(* IEC 61131-3 sources: daoli-st-library/DL_Device (part 21) *)

(* ---- FB_DL_EscChuckCurrentMonitor.st ---- *)
(*
    FB_DL_EscChuckCurrentMonitor —— ESC 静电吸附电流监视
    ------------------------------------------------------------------
    分类      : DL_Device / Diagnostics
    前缀      : FB_DL_
    版本      : 1.0.0
    溯源      : 半导体静电吸盘（ESC）自研线，clean-room 自研，无可挖开源源；
                只借公开半导体设备工程语义（吸附/建立/稳态/释放三段，失吸与打火是
                可区分的失效模式）；判据、状态机、错误分级与码位 100% 自有；
                E_DL_Ne107Status 属主为 I_DL_DeviceHealth，本件只引用不重声明（R70）
    平台      : 纯 IEC 61131-3，CODESYS V3.5+ / TwinCAT 3 / InoProShop 通用
    作者      : 道莅代码库 · PLC编程专家（R19）
    ------------------------------------------------------------------
    功能说明  : 吸附电压施加后电流须在 tBuildTime 内落进电流窗（建立段）；之后电流须
                持续落窗（稳态段，低于下限超 tConfirmTime 判失吸）；撤电压后电流须归零
                （释放段）。失吸会导致晶圆飞片/破片，打火会烧盘面，两者在电流波形上
                是两种截然不同的特征，本件把「电流长时间偏低」与「瞬时尖峰」分开判。
                核心防御：① 阈值倒置先自动交换并置信息码，交换后仍非法才报故障级；
                ② 电流/电压非有限即故障级并冻结判定，且保持末次 bAttached——
                   把正在吸附的晶圆判成飞片会引发误停机；
                ③ 电压低于吸附门限时不判电流（电压没加上，电流当然为零），回 eIdle；
                ④ 打火只锁存并出口 eOutOfSpec，不置 bError（可继续生产但需检修）；
                ⑤ 泄漏趋势用前后半窗均值比较，只置信息级不置故障。
                职责边界：吸附电压给定与放电归静电电源件，本件只判电流形态。
    错误码    : 16#0003_016E 电流窗上下限倒置已自动交换 / 泄漏趋势上升 / 贴近边界降级运行——信息级，正常防御
                16#0003_016F 预留禁用（信息级，不得挪用）
                16#0003_0336 阈值参数非法或输入非有限——故障级，判定冻结且保持末次吸附结论
                16#0003_0337 建立超时或稳态电流失窗（判失吸）——故障级，eHealth = eFailure
                16#0003_0338 打火尖峰锁存——故障级码位且 eHealth = eOutOfSpec，但按 R13 家族裁定不置 bError
    码位总账  : 16#0003_016E 用 / 16#0003_016F 预留 ｜ 16#0003_0336 用 / 16#0003_0337 用 / 16#0003_0338 用
    状态机    : E_DL_EscState（eIdle / eBuild / eSteady / eRelease / eFault）五态，CASE 含 ELSE 兜底，
                ELSE 回 eFault 并置故障级 0336。
    采样约定  : fbTrigReset / fbBuild / fbLossConfirm 在本体首部无条件刷新——两个定时器的 IN
                由状态导出但调用绝不放进 IF 或 CASE（按段断输入是本族高危点）；
                采样周期越域即故障级，因为趋势窗与确认时间都隐含依赖采样节拍。
    修订记录  : 2026-11-16 v1.0.0 首次入库（R19）
*)

(*
    枚举 : E_DL_EscState —— 静电吸盘工作段（本文件为全库唯一属主）
*)
TYPE E_DL_EscState :
(
    eIdle    := 0,                            // 空闲：未施加吸附电压 / idle, no chuck voltage applied
    eBuild   := 1,                            // 建立段：等待电流落窗 / build phase, waiting for the current to settle
    eSteady  := 2,                            // 稳态段：电流持续落窗 / steady phase, the current stays inside the window
    eRelease := 3,                            // 释放段：等待电流归零 / release phase, waiting for the current to vanish
    eFault   := 4                             // 故障：判定冻结 / fault, evaluation frozen
);
END_TYPE

FUNCTION_BLOCK FB_DL_EscChuckCurrentMonitor
VAR_INPUT
    bEnable         : BOOL;                   // 使能，FALSE 撤销所有判定输出 / enable, FALSE withdraws every judgement output
    bReset          : BOOL;                   // 复位，上升沿清故障与趋势 / reset, rising edge clears the faults and the trend
    bChuckOn        : BOOL := FALSE;          // 吸附电压施加命令（上层给定）/ chuck voltage command from the upper layer
    fChuckCurrent   : REAL := 0.0;            // 吸附电流测量值 [uA]，范围 0.0~10000.0 / chuck current measurement [uA], range 0.0~10000.0
    fChuckVoltage   : REAL := 0.0;            // 吸附电压测量值 [V]，范围 0.0~5000.0 / chuck voltage measurement [V], range 0.0~5000.0
    fCurMin         : REAL := 5.0;            // 稳态电流窗下限 [uA]，必须 > 0 / steady window lower bound [uA], must be > 0
    fCurMax         : REAL := 500.0;          // 稳态电流窗上限 [uA]，必须 > fCurMin / steady window upper bound [uA], must be > fCurMin
    fSparkRise      : REAL := 50.0;           // 打火判据：单拍电流跳变量阈值 [uA]，必须 > 0 / spark criterion, per cycle current step [uA], must be > 0
    tBuildTime      : TIME := T#2S;           // 建立段允许时长 [ms]，范围 100~30000 / build phase allowance [ms], range 100~30000
    tConfirmTime    : TIME := T#500MS;        // 失吸确认时间 [ms]，范围 0~10000 / loss confirmation time [ms], range 0~10000
    tSampleTime     : TIME := T#10MS;         // 采样周期 [ms]，范围 1~1000 / sample time [ms], range 1~1000
END_VAR
VAR_OUTPUT
    bAttached       : BOOL;                   // 判定已吸附（建立成功且稳态落窗）/ attached, build succeeded and the steady current stays in the window
    bSpark          : BOOL;                   // 检出打火尖峰（锁存）/ spark peak detected, latched
    bLeakTrend      : BOOL;                   // 泄漏趋势上升（盘面污染或绝缘退化）/ leakage trend rising, contamination or insulation ageing
    bDegraded       : BOOL;                   // 降级运行（电流在窗内但贴近边界）/ degraded, the current is in the window but close to a bound
    eHealth         : E_DL_Ne107Status;       // 健康出口（引用唯一属主枚举）/ health output referencing the owner enumeration
    uAttachCount    : UDINT;                  // 累计成功吸附次数，饱和 [次] / accumulated successful attaches, saturating [times]
    eErr            : UDINT;                  // 错误码，0=正常 / error id, 0=ok
    bError          : BOOL;                   // 故障标志，eErr 为故障级时 TRUE / error flag, TRUE on fault-level eErr
END_VAR
VAR
    eState          : E_DL_EscState := eIdle; // 状态机当前态 / current state machine state
    fbTrigReset     : R_TRIG;                 // 复位上升沿实例，本体首部无条件刷新 / reset edge instance, refreshed unconditionally
    fbBuild         : TON;                    // 建立段定时器，本体首部无条件刷新 / build phase timer, refreshed unconditionally
    fbLossConfirm   : TON;                    // 失吸确认定时器，本体首部无条件刷新 / loss confirmation timer, refreshed unconditionally
    fPrevCur        : REAL;                   // 上一拍电流，用于打火跳变判据 [uA] / previous current for the spark step test [uA]
    fTrendAcc       : REAL;                   // 后窗电流均值累加 [uA] / second window current mean accumulator [uA]
    fTrendBase      : REAL;                   // 前窗电流均值累加 [uA] / first window current mean accumulator [uA]
    uTrendCnt       : UINT;                   // 趋势取样计数 [拍] / trend sampling counter [scan]
    fCurMinEff      : REAL;                   // 交换与钳位后的电流窗下限 [uA] / effective lower bound after swap and clamp [uA]
    fCurMaxEff      : REAL;                   // 交换与钳位后的电流窗上限 [uA] / effective upper bound after swap and clamp [uA]
    fBandEff        : REAL;                   // 近边界判定带宽 [uA] / near boundary band width [uA]
    fCur            : REAL;                   // 本拍电流副本 [uA] / current copy of this cycle [uA]
    bNonFin         : BOOL;                   // 输入非有限判定标志 / non-finite input flag
    bInWindow       : BOOL;                   // 电流落窗判定 / current inside the window
    bInit           : BOOL := FALSE;          // 首扫标志，初值 FALSE，判据 NOT bInit / first-scan flag, initial FALSE, tested with NOT
END_VAR
VAR CONSTANT
    DL_ESC_CUR_ABS_MAX : REAL := 10000.0;     // 电流绝对上限（三阈值钳位用）[uA] / absolute current bound used by the clamps [uA]
    DL_ESC_VOLT_MIN    : REAL := 100.0;       // 判定「电压确实加上了」的下限 [V] / lower bound proving the voltage is really applied [V]
    DL_ESC_TREND_N     : UINT := 50;          // 趋势取样个数 [拍] / number of trend samples [scan]
    DL_ESC_BAND_RATIO  : REAL := 0.05;        // 近边界判定带宽（相对窗宽）[无量纲] / near boundary band relative to the window [dimensionless]
    DL_ESC_DT_MAX      : TIME := T#1S;        // 采样周期上限 [ms] / sample time upper bound [ms]
    DL_ESC_DT_MIN      : TIME := T#1MS;       // 采样周期下限 [ms] / sample time lower bound [ms]
    DL_FLOAT_EPS       : REAL := 1.0E-6;      // 浮点判等容差 [无量纲] / float equality tolerance [dimensionless]
    DL_ESC_TWO         : REAL := 2.0;         // 二值常量，窗口折半用 [无量纲] / two, used to halve the trend window
    DL_ESC_INF_GUARD   : REAL := 1.0E38;      // 非有限幅值判定阈值 [无量纲] / non-finite magnitude guard [dimensionless]
    DL_ESC_CNT_MAX     : UDINT := 16#FFFF_FFFE; // 吸附计数饱和值 [次] / attach counter saturation value [times]
    DL_ESC_ZERO        : REAL := 0.0;         // 零值常量，避免裸字面量 [无量纲] / zero constant, avoids a bare literal [dimensionless]
END_VAR

// 段 1｜边沿与定时器实例无条件周期刷新（红线：严禁放入条件分支）/ segment 1, unconditional refresh
fbTrigReset(CLK := bReset);
fbBuild(IN := (eState = eBuild) AND bEnable, PT := tBuildTime); // 仅建立段计时 / the timer runs only during the build phase
fbLossConfirm(IN := (eState = eSteady) AND bEnable AND (fChuckCurrent < fCurMin), PT := tConfirmTime); // 仅稳态且电流低于下限时计时 / runs only in the steady phase while the current is below the bound

// 段 2｜输出与错误状态预置（bAttached / bSpark 为保持量，不预置）/ segment 2, preset outputs, the held flags are not preset
eErr := 0;                                    // 预置无错误 / preset no error
bError := FALSE;                              // 预置无故障 / preset no fault
bDegraded := FALSE;                           // 预置未降级 / preset not degraded
bLeakTrend := FALSE;                          // 预置无泄漏趋势 / preset no leakage trend
eHealth := eOk;                               // 预置健康 / preset OK

// 段 3｜首扫初始化（唯一合法范式：初值 FALSE，判据 NOT bInit）/ segment 3, first-scan initialisation
IF NOT bInit THEN
    bAttached := FALSE;                       // 首扫不判吸附 / no attach survives the first scan
    bSpark := FALSE;                          // 首扫不打火锁存 / no spark latch survives the first scan
    uAttachCount := 0;                        // 吸附计数清零 / clear the attach counter
    fPrevCur := fChuckCurrent;                // 电流基准取当前测量，避免首拍误判打火 / seed the current reference to avoid a false spark on the first scan
    uTrendCnt := 0;                          // 趋势计数清零 / clear the trend counter
    fTrendAcc := DL_ESC_ZERO;                 // 后窗累加清零 / clear the second window accumulator
    fTrendBase := DL_ESC_ZERO;                // 前窗累加清零 / clear the first window accumulator
    bInit := TRUE;                            // 首扫只做一次 / first scan runs once only
END_IF

// 段 4｜使能闸：失能撤销全部判定输出 / segment 4, enable gate
IF NOT bEnable THEN
    bAttached := FALSE;                       // 撤销吸附判定 / withdraw the attach judgement
    bDegraded := FALSE;                       // 撤销降级 / withdraw the degraded flag
    bLeakTrend := FALSE;                      // 撤销趋势 / withdraw the trend flag
    eHealth := eUnknown;                      // 失能即未知 / unknown while disabled
    RETURN;                                   // 失能即出口 / disabled is the exit
END_IF

// 段 5｜阈值交换与合法性闸（倒置先交换，交换后仍非法才报故障）/ segment 5, threshold swap and validity
fCurMinEff := fCurMin;                        // 取入参副本 / copy the input
fCurMaxEff := fCurMax;                        // 取入参副本 / copy the input
IF fCurMaxEff < fCurMinEff THEN
    fCurMinEff := fCurMax;                    // 交换：下限取原上限 / swap, the lower bound takes the former upper bound
    fCurMaxEff := fCurMin;                    // 交换：上限取原下限 / swap, the upper bound takes the former lower bound
    eErr := 16#0003_016E;                     // 信息级：上下限倒置已自动交换 / info level, the inverted bounds were swapped
END_IF
fCurMinEff := MIN(MAX(fCurMinEff, DL_ESC_ZERO), DL_ESC_CUR_ABS_MAX); // 下限收敛到物理域 / converge the lower bound into the physical domain
fCurMaxEff := MIN(MAX(fCurMaxEff, DL_ESC_ZERO), DL_ESC_CUR_ABS_MAX); // 上限收敛到物理域 / converge the upper bound into the physical domain
IF (fCurMinEff <= DL_FLOAT_EPS) OR (fCurMaxEff <= fCurMinEff) THEN
    eErr := 16#0003_0336;                     // 阈值非法故障码 / illegal threshold fault id
    bError := TRUE;                           // 置故障标志 / raise the error flag
    eState := eFault;                         // 落故障态，判定冻结 / enter the fault state, the evaluation is frozen
    eHealth := eFailure;                      // 阈值不可信即出口失效 / untrustworthy thresholds mean a failed health output
    RETURN;                                   // 故障级提前返回，bAttached 保持末值 / early return, bAttached keeps its last value
END_IF
fBandEff := DL_ESC_BAND_RATIO * (fCurMaxEff - fCurMinEff); // 近边界带宽 [uA] / near boundary band width [uA]

// 段 6｜输入非有限闸：冻结判定并保持末次吸附结论 / segment 6, non-finite gate freezes the judgement
bNonFin := (fChuckCurrent <> fChuckCurrent) OR (fChuckCurrent > DL_ESC_INF_GUARD) OR (fChuckCurrent < -DL_ESC_INF_GUARD)
        OR (fChuckVoltage <> fChuckVoltage) OR (fChuckVoltage > DL_ESC_INF_GUARD) OR (fChuckVoltage < -DL_ESC_INF_GUARD)
        OR (fSparkRise <> fSparkRise);        // 非有限判定 / non-finite detection
IF bNonFin THEN
    eErr := 16#0003_0336;                     // 输入非有限故障码 / non-finite input fault id
    bError := TRUE;                           // 置故障标志 / raise the error flag
    eState := eFault;                         // 落故障态 / enter the fault state
    eHealth := eFailure;                      // 测量不可信 / the measurement is untrustworthy
    RETURN;                                   // 保持末次 bAttached，绝不掉成未吸附 / keep the last attach state, never fall back to detached
END_IF

// 段 7｜采样周期闸（趋势窗与确认时间都依赖采样节拍）/ segment 7, sample time gate
IF (tSampleTime < DL_ESC_DT_MIN) OR (tSampleTime > DL_ESC_DT_MAX) THEN
    eErr := 16#0003_0336;                     // 采样周期非法故障码 / illegal sample time fault id
    bError := TRUE;                           // 置故障标志 / raise the error flag
    eState := eFault;                         // 落故障态 / enter the fault state
    eHealth := eFailure;                      // 节拍不可信 / the timing is untrustworthy
    RETURN;                                   // 出口 / exit
END_IF

// 段 8｜复位沿清故障与趋势（不改变已建立的吸附结论）/ segment 8, reset clears the faults and the trend
IF fbTrigReset.Q THEN
    bSpark := FALSE;                          // 清打火锁存 / clear the spark latch
    bLeakTrend := FALSE;                      // 清趋势 / clear the trend
    uTrendCnt := 0;                           // 清趋势计数 / clear the trend counter
    fTrendAcc := DL_ESC_ZERO;                 // 清后窗累加 / clear the second window
    fTrendBase := DL_ESC_ZERO;                // 清前窗累加 / clear the first window
    IF eState = eFault THEN
        eState := eIdle;                      // 故障态复位回空闲 / a reset leaves the fault state
    END_IF
END_IF

// 段 9｜电流副本与落窗判定 / segment 9, current copy and window test
fCur := fChuckCurrent;                        // 取入参副本 [uA] / copy the input [uA]
bInWindow := (fCur >= fCurMinEff) AND (fCur <= fCurMaxEff); // 落窗判定 / window test

// 段 10｜打火判据（单拍跳变 + 吸附电压在场，只锁存不置 bError）/ segment 10, spark criterion
IF bChuckOn AND (ABS(fCur - fPrevCur) > fSparkRise) THEN
    bSpark := TRUE;                           // 锁存打火 / latch the spark
    eErr := 16#0003_0338;                     // 打火故障级码位，但按家族裁定不置 bError / spark fault id without raising bError
    eHealth := eOutOfSpec;                    // 能继续吸不等于盘面完好 / still holding does not mean the chuck surface is intact
END_IF
fPrevCur := fCur;                             // 记录本拍电流供下一拍比较 / remember this cycle current

// 段 11｜降级判定：电流在窗内但贴近上下边界 / segment 11, degraded evaluation near a bound
IF bInWindow AND ((fCur <= (fCurMinEff + fBandEff)) OR (fCur >= (fCurMaxEff - fBandEff))) THEN
    bDegraded := TRUE;                        // 贴近边界即降级 / closeness to a bound is a degradation
    IF eErr = 0 THEN
        eErr := 16#0003_016E;                 // 信息级：贴近边界降级运行 / info level, running degraded near a bound
    END_IF
END_IF

// 段 12｜泄漏趋势（前后半窗均值比较，只置信息级）/ segment 12, leakage trend by half window means
IF eState = eSteady THEN
    IF uTrendCnt < (DL_ESC_TREND_N / 2) THEN
        fTrendBase := fTrendBase + fCur / (UINT_TO_REAL(DL_ESC_TREND_N) / DL_ESC_TWO); // 前窗均值累加 [uA] / accumulate the first window mean [uA]
        uTrendCnt := uTrendCnt + 1;           // 计数加一 / increment the counter
    ELSE
        fTrendAcc := fTrendAcc + fCur / (UINT_TO_REAL(DL_ESC_TREND_N) / DL_ESC_TWO);   // 后窗均值累加 [uA] / accumulate the second window mean [uA]
        uTrendCnt := uTrendCnt + 1;           // 计数加一 / increment the counter
        IF uTrendCnt >= DL_ESC_TREND_N THEN
            IF fTrendAcc > (fTrendBase + DL_ESC_BAND_RATIO * (fCurMaxEff - fCurMinEff)) THEN
                bLeakTrend := TRUE;           // 后窗显著上爬：污染或绝缘退化 / the second window creeps up, contamination or insulation ageing
                eErr := 16#0003_016E;         // 信息级：泄漏趋势上升 / info level, the leakage trend is rising
                eHealth := eMaintenanceReq;   // 需安排检修 / maintenance is required
            END_IF
            uTrendCnt := 0;                   // 窗口滑动复位 / restart the sliding window
            fTrendAcc := DL_ESC_ZERO;         // 后窗累加清零 / clear the second window
            fTrendBase := DL_ESC_ZERO;        // 前窗累加清零 / clear the first window
        END_IF
    END_IF
END_IF

// 段 13｜状态机（含 ELSE 兜底）/ segment 13, state machine with ELSE fallback
CASE eState OF
    eIdle:
        bAttached := FALSE;                   // 空闲即未吸附 / idle means detached
        IF bChuckOn AND (fChuckVoltage >= DL_ESC_VOLT_MIN) THEN
            eState := eBuild;                 // 电压确实加上才进入建立段 / enter the build phase only when the voltage is really present
        END_IF

    eBuild:
        IF bInWindow THEN
            eState := eSteady;                // 电流落窗即建立成功 / the current entering the window completes the build
            bAttached := TRUE;                // 判定已吸附 / mark it attached
            IF uAttachCount < DL_ESC_CNT_MAX THEN
                uAttachCount := uAttachCount + 1; // 饱和计数 / saturating count
            END_IF
        ELSIF fbBuild.Q THEN
            eErr := 16#0003_0337;             // 建立超时故障码 / build timeout fault id
            bError := TRUE;                   // 置故障标志 / raise the error flag
            eHealth := eFailure;              // 失吸 / the wafer is not held
            eState := eFault;                 // 落故障态 / enter the fault state
            bAttached := FALSE;               // 建立失败即未吸附 / a failed build means detached
        END_IF

    eSteady:
        bAttached := TRUE;                    // 稳态保持吸附 / the steady phase keeps the attach state
        IF NOT bChuckOn THEN
            eState := eRelease;               // 撤电压即进入释放段 / releasing the voltage enters the release phase
        ELSIF fbLossConfirm.Q THEN
            eErr := 16#0003_0337;             // 失吸确认故障码 / loss confirmation fault id
            bError := TRUE;                   // 置故障标志 / raise the error flag
            eHealth := eFailure;              // 失吸 / the wafer is lost
            eState := eFault;                 // 落故障态 / enter the fault state
            bAttached := FALSE;               // 确认失吸 / confirmed detached
        END_IF

    eRelease:
        bAttached := FALSE;                   // 释放段即不再算吸附 / the release phase is not an attached state
        IF fCur <= DL_FLOAT_EPS THEN
            eState := eIdle;                  // 电流归零即回空闲 / back to idle once the current vanishes
        ELSIF bChuckOn THEN
            eState := eBuild;                 // 释放过程中重新上电：重新建立 / re-energising during release restarts the build
        END_IF

    eFault:
        bAttached := FALSE;                   // 故障态不判吸附 / no attach judgement in the fault state
        IF NOT bChuckOn THEN
            eState := eIdle;                  // 撤电压允许退出故障态（复位亦可）/ withdrawing the voltage also leaves the fault state
        END_IF

ELSE
    eErr := 16#0003_0336;                     // 故障级：非法状态兜底 / fault level, illegal state fallback
    bError := TRUE;                           // 置故障标志 / raise the error flag
    eState := eFault;                         // 回故障态 / fall back to the fault state
    eHealth := eUnknown;                      // 状态不可信 / the state is untrustworthy
END_CASE
END_FUNCTION_BLOCK

(* ---- FB_DL_EsdGroundMonitor.st ---- *)
(*
  ==================================================================
  组件名 Component  : FB_DL_EsdGroundMonitor
  分类   Category   : DL_Device
  复杂度 Complexity  : cx4
  版本   Version    : 1.0.0
  功能   Purpose    : ESD 接地连续性监视。对接地电阻做窗口判级（低于下限疑短路 /
                      接线反，高于上限疑断路），双阈值迟滞防边界抖动；传感失效
                      锁存优先于判级；健康语言出口按 NE107 五态口径输出。
  来源   Source     : self-esc（次源 t2-8 NE107，借鉴 NE107 健康状态五态语言，
                      clean-room 自研实现，未复制任何文档代码行）
  溯源   Origin     : IEC 61131-3 标准语义的道莅防御性实现；ESD 接地电阻窗口
                      判级为公开防静电工艺语义（常见口径 <10 欧姆量级）。
  平台   Platform   : 纯 IEC 61131-3（LREAL 运算，无私有库、无定时器实例）
  分工声明 Split     : 与 DL_Device 存量联锁族（风机关 / 传递窗）分工——本件只
                      做接地电阻判级与健康语言映射，不做风量联锁与顺控。
  作者   Author     : 道莅代码库 · PLC 编程专家（R57）
  ------------------------------------------------------------------
  边界 Boundary     :
                      一 组态闸（R151）：fOhmMin > 0 且 fOhmMax > fOhmMin，
                         迟滞带宽 0 <= fHystOhm < 半窗宽；
                      二 迟滞收窄口径：进入判据用全带宽，退出判据带宽收窄
                         fHystOhm，防边界抖动反复置清；
                      三 传感失效（非有限双判据 / 电阻 < 0）锁存优先于判级；
                      四 成因锁存解除路径 = bReset 上升沿（唯一路径，R188）；
                      五 无全局变量、无外部变量声明、无物理地址寻址。
  输出契约 Output contract:
                      eHealth 为 NE107 五态健康语言；bGroundOk 为放行派生电平；
                      eFault 为锁存回放；bError 与故障级成因配对（R45）。
  修订记录 Revision  :
    2026-11-21  v1.0.0  R57 首版（批 4 · 序号 16）
  ==================================================================
*)

TYPE E_DL_EgmPhase :
(
    eIdle  := 0,  // 未使能：判级停摆 / disabled, the grading idle
    eRun   := 10, // 运行：逐拍判级 / running, graded every scan
    eFault := 90  // 故障：成因锁存 / fault, the cause latched
);
END_TYPE

TYPE E_DL_EgmFault :
(
    eNone       := 0, // 无成因 / no cause
    eCfgIllegal := 1, // 组态非法：电阻窗或迟滞越域（故障级，与 bError 配对）/ an illegal config
    eSensorBad  := 2, // 传感失效：电阻非有限或负值（故障级，与 bError 配对）/ a sensor failure
    eGroundOpen := 3, // 接地断路：电阻超上限（故障级，与 bError 配对）/ a ground open
    eGroundShort:= 4, // 接地短路疑点：电阻低于下限（故障级，与 bError 配对）/ a ground short suspect
    ePhaseBad   := 5  // 非法相位兜底（故障级，与 bError 配对）/ an illegal phase fallback
);
END_TYPE

TYPE E_DL_EgmHealth :
(
    eInit           := 0, // NE107 初始态 / the NE107 initial state
    eGood           := 1, // NE107 正常 / the NE107 good state
    eCheckFunction  := 2, // NE107 功能受影响（组态非法驻留）/ the NE107 check function state
    eMaintenanceReq := 3, // NE107 维护要求（判级异常驻留）/ the NE107 maintenance required state
    eFailure        := 4  // NE107 故障（传感失效锁存）/ the NE107 failure state
);
END_TYPE

FUNCTION_BLOCK FB_DL_EsdGroundMonitor
VAR_INPUT
    bEnable   : BOOL := TRUE;   // 使能，失能时判级停摆 [-] / enable, the grading stops when disabled
    bReset    : BOOL := FALSE;  // 复位上升沿清全部成因锁存 [-] / reset rising edge clears every cause latch
    fResOhm   : LREAL := 5.0;   // 接地电阻实测 [欧姆] / the measured ground resistance [ohm]
    fOhmMin   : LREAL := 0.5;   // 电阻窗下限 [欧姆]，域 大于零 / the window floor [ohm], above zero
    fOhmMax   : LREAL := 10.0;  // 电阻窗上限 [欧姆]，域 大于下限 / the window ceiling [ohm], above the floor
    fHystOhm  : LREAL := 0.5;   // 迟滞带宽 [欧姆]，域 0..半窗宽 / the hysteresis band [ohm]
END_VAR
VAR_OUTPUT
    eHealth  : E_DL_EgmHealth := E_DL_EgmHealth.eInit; // NE107 健康语言出口 [枚举] / the NE107 health outlet [enum]
    bGroundOk: BOOL := FALSE; // 接地合格放行派生电平 [-] / the ground ok derived level
    ePhase   : E_DL_EgmPhase := E_DL_EgmPhase.eIdle; // 相位出口 [枚举] / the phase outlet [enum]
    eFault   : E_DL_EgmFault := E_DL_EgmFault.eNone; // 成因出口，锁存回放 [枚举] / the cause outlet replayed from the latch
    bError   : BOOL := FALSE; // 故障锁存标志 [-] / the fault latch flag
END_VAR
VAR
    rtReset : R_TRIG; // 复位沿检测，段 0 无条件刷新 / the reset edge, refreshed unconditionally
    _ePhase : E_DL_EgmPhase := E_DL_EgmPhase.eIdle; // 内部相位，CASE 唯一写入目标 / the internal phase
    _eFaulC : E_DL_EgmFault := E_DL_EgmFault.eNone; // 故障级成因，锁存至复位沿 / the fault cause, latched until the reset edge
    _bFault : BOOL := FALSE; // 故障锁存位 [-] / the fault latch bit
    _bInit  : BOOL := FALSE; // 首扫初始化完成标志（R310）/ the first scan flag
    _bInOk  : BOOL := FALSE; // 电阻有限且非负 [-] / the resistance finite and nonnegative
    _bCfgOk : BOOL := FALSE; // 组态域内 [-] / the configuration inside the domain
    _bOpen  : BOOL := FALSE; // 断路迟滞锁存 [-] / the open hysteresis latch
    _bShort : BOOL := FALSE; // 短路疑点迟滞锁存 [-] / the short suspect hysteresis latch
END_VAR

// 段 0｜沿检测无条件周期刷新（禁入分支）/ segment 0, the unconditional refresh
rtReset(CLK := bReset); // 复位沿 / the reset edge

// 段 1｜首扫初始化（R310）/ segment 1, the first scan initialisation
IF NOT _bInit THEN // 首扫一拍 / the first scan
    _bInit  := TRUE; // 置首扫标志 / raise the flag
    _ePhase := E_DL_EgmPhase.eRun; // 相位从运行起步（使能默认真）/ the phase starts in run
END_IF

// 段 2｜复位沿作用域：清锁存 / 清迟滞 / 迁相位（三项逐项声明）/ segment 2, the reset edge scope
IF rtReset.Q THEN // 复位沿 / the reset edge
    _bFault := FALSE; // 作用域一：清故障锁存 / scope one, clear the fault latch
    _eFaulC := E_DL_EgmFault.eNone; // 作用域一：清成因 / scope one, clear the cause
    _bOpen := FALSE; // 作用域二：清断路迟滞 / scope two, clear the open latch
    _bShort := FALSE; // 作用域二：清短路迟滞 / scope two, clear the short latch
    _ePhase := E_DL_EgmPhase.eRun; // 作用域三：迁回运行相 / scope three, back to run
END_IF

// 段 3｜组态与输入域闸（R151 全覆盖，边界一）/ segment 3, the configuration and input gates
_bInOk := (fResOhm = fResOhm) AND ((fResOhm - fResOhm) = (fResOhm - fResOhm)) AND (fResOhm >= 0.0); // 电阻有限且非负 / the resistance finite and nonnegative
_bCfgOk := (fOhmMin > 0.0) AND (fOhmMin = fOhmMin) AND (fOhmMax > fOhmMin) AND (fOhmMax = fOhmMax) AND (fHystOhm >= 0.0) AND (fHystOhm < (fOhmMax - fOhmMin) / 2.0); // 窗与迟滞域判定（除子为窗宽已证大于零）/ the window and hysteresis verdict
IF (NOT _bInOk) OR (NOT _bCfgOk) THEN // 输入缺陷或组态非法 / an input defect or an illegal config
    IF NOT _bFault THEN // 未锁存才迁移（防同拍抹除）/ migrate only while unlatched
        _bFault := TRUE; // 置故障锁存 / raise the fault latch
        IF NOT _bInOk THEN // 传感失效优先归因（R190 归因唯一）/ the sensor failure attributed first
            _eFaulC := E_DL_EgmFault.eSensorBad; // 传感失效成因 / the sensor cause
        ELSE // 组态非法 / the illegal config
            _eFaulC := E_DL_EgmFault.eCfgIllegal; // 组态成因 / the config cause
        END_IF
        _ePhase := E_DL_EgmPhase.eFault; // 迁故障相 / migrate to fault
    END_IF
END_IF

// 段 4｜相位机：ENUM + CASE，含 ELSE 非法相位兜底（R128）/ segment 4, the phase machine
CASE _ePhase OF

E_DL_EgmPhase.eIdle: // 未使能相：健康语言回初始 / the idle phase, the health back to init
    IF bEnable AND (NOT _bFault) THEN // 使能且无故障 / enabled and unfaulted
        _ePhase := E_DL_EgmPhase.eRun; // 迁运行相 / migrate to run
    END_IF

E_DL_EgmPhase.eRun: // 运行相：逐拍判级 / the run phase, graded every scan
    IF NOT bEnable THEN // 失能 / disabled
        _ePhase := E_DL_EgmPhase.eIdle; // 迁未使能相 / migrate to idle
    ELSE // 正常判级 / the normal grading
        IF fResOhm > fOhmMax THEN // 断路进入判据（全带宽）/ the open entry criterion, the full band
            _bOpen := TRUE; // 置断路迟滞 / raise the open latch
        ELSIF fResOhm < fOhmMax - fHystOhm THEN // 断路退出判据（迟滞收窄，边界二）/ the open exit criterion, the narrowed band
            _bOpen := FALSE; // 清断路迟滞 / clear the open latch
        END_IF
        IF fResOhm < fOhmMin THEN // 短路疑点进入判据（全带宽）/ the short entry criterion
            _bShort := TRUE; // 置短路迟滞 / raise the short latch
        ELSIF fResOhm > fOhmMin + fHystOhm THEN // 短路退出判据（迟滞收窄）/ the short exit criterion
            _bShort := FALSE; // 清短路迟滞 / clear the short latch
        END_IF
        IF _bShort THEN // 短路疑点优先（接线异常更急）/ the short suspect first
            _bFault := TRUE; // 置故障锁存 / raise the fault latch
            _eFaulC := E_DL_EgmFault.eGroundShort; // 故障级成因（R45 配对 bError）/ the fault cause
            _ePhase := E_DL_EgmPhase.eFault; // 迁故障相 / migrate to fault
        ELSIF _bOpen THEN // 断路次优先 / the open next
            _bFault := TRUE; // 置故障锁存 / raise the fault latch
            _eFaulC := E_DL_EgmFault.eGroundOpen; // 故障级成因（R45 配对 bError）/ the fault cause
            _ePhase := E_DL_EgmPhase.eFault; // 迁故障相 / migrate to fault
        END_IF
    END_IF

E_DL_EgmPhase.eFault: // 故障相：成因锁存，等待复位沿；健康语言按成因映射 / the fault phase, the cause latched until the reset edge

ELSE // 非法相位兜底（R128）/ the illegal phase fallback
    _bFault := TRUE; // 置故障锁存 / raise the fault latch
    _eFaulC := E_DL_EgmFault.ePhaseBad; // 故障级成因（R45 配对 bError）/ the fault cause
    _ePhase := E_DL_EgmPhase.eFault; // 迁故障相 / migrate to fault
END_CASE

// 段 5｜统一出口：健康语言与放行派生单点映射 / segment 5, the unified outlet
IF _bFault THEN // 故障锁存优先 / the fault latch first
    eFault := _eFaulC; // 成因锁存回放（R152）/ the cause replayed
    CASE _eFaulC OF // 成因到 NE107 健康语言映射 / the cause to health mapping
    E_DL_EgmFault.eSensorBad: eHealth := E_DL_EgmHealth.eFailure; // 传感失效映射故障态 / the sensor failure to failure
    E_DL_EgmFault.eCfgIllegal: eHealth := E_DL_EgmHealth.eCheckFunction; // 组态非法映射功能受影响 / the config to check function
    ELSE eHealth := E_DL_EgmHealth.eMaintenanceReq; // 判级异常映射维护要求 / the grading anomalies to maintenance
    END_CASE
ELSE // 无锁存 / no latch
    eFault := E_DL_EgmFault.eNone; // 无成因 / no cause
    IF bEnable THEN // 使能中 / enabled
        eHealth := E_DL_EgmHealth.eGood; // 健康态 / the good state
    ELSE // 失能驻留 / disabled
        eHealth := E_DL_EgmHealth.eInit; // 初始态 / the init state
    END_IF
END_IF
bGroundOk := (_ePhase = E_DL_EgmPhase.eRun) AND (NOT _bFault) AND (NOT _bShort) AND (NOT _bOpen); // 放行派生电平 / the ok derived level
ePhase := _ePhase; // 相位出口单点映射 / the phase outlet
bError := _bFault; // 故障标志与锁存位同源 / the flag shares the latch
END_FUNCTION_BLOCK

(* ---- FB_DL_ExhaustDpTrend.st ---- *)
(*
  FB_DL_ExhaustDpTrend  —  尾气管路压差趋势监视与堵塞预警 / Exhaust line differential-pressure trend and clog warning
  分类 Category : DL_Device
  码位 Code     : 16#03_2_08
  版本 Version  : 1.0.0
  溯源 Source   : LGF Measurement 语义借鉴 · clean-room 实现，仅借分类/参数域/命名，未复制源码
  功能 Function : 1) 尾气前后压差滑动窗统计（复用 FB_DL_SignalStatistics）；
                  2) 周期末均值快照对比折算趋势 [kPa/天]；
                  3) 堵塞预警分级（预警级带迟滞，严重级持续确认升级）。
  边界 Boundary : ① 风机停机时冻结趋势累计（禁把停机零流量当堵塞）；
                  ② 压差无效剔除并置掩码；
                  ③ 趋势窗样本不足不出结论；
                  ④ 预警阈值带迟滞且解除可达；
                  ⑤ 输出三行同向：压差均值 → 趋势斜率 → 堵塞预警。
  依赖 Depends  : FB_DL_SignalStatistics × 2（当前窗 / 快照窗，每拍无条件调用）

  码表 Error codes（本件子码步进 16#10，避让邻件码位）:
    16#0002_0308 故障级：组态非法（周期/门限/迟滞 <= 0）
    16#0002_0318 故障级：严重堵塞（压差持续超严重门限，锁存需复位）
    16#0002_0328 信息级：压差无效剔除 / 样本不足不出结论 / 风机停机趋势冻结（不置 bError）
*)

TYPE E_DL_ExtPhase :
(
    eIdle  := 0,  // 空闲 / Idle
    eWatch := 10, // 压差趋势监视 / DP trend watching
    eFault := 90  // 组态故障锁定 / Configuration fault locked
);
END_TYPE

FUNCTION_BLOCK FB_DL_ExhaustDpTrend
VAR_INPUT
    bEnable       : BOOL;                           // 总使能，FALSE 回空闲 / Master enable
    bReset        : BOOL;                           // 复位，上升沿清故障 / Reset, clears fault
    fDpKpa        : REAL;                           // 尾气前后压差 [kPa] / Exhaust differential pressure [kPa]
    bFanRunning   : BOOL;                           // 风机运行反馈 / Fan running feedback
    uPeriodMin    : UINT := 60;                     // 趋势统计周期 [min]，域 > 0 / Trend period [min]
    fWarnKpa      : REAL := 2.5;                    // 堵塞预警门限 [kPa] / Clog warning threshold [kPa]
    fTripKpa      : REAL := 4.0;                    // 严重堵塞门限 [kPa] / Severe clog threshold [kPa]
    fHystKpa      : REAL := 0.3;                    // 预警迟滞 [kPa]，域 > 0 / Warning hysteresis [kPa]
    uTripConfirm  : UINT := 10;                     // 严重堵塞确认拍数 [拍] / Severe confirm scans
    fTaskCycle    : REAL := 1.0;                    // 任务周期 [s]，域 > 0 / Task cycle [s]
    fEps          : REAL := 1.0E-6;                 // 浮点判零容差 [1] / Floating zero tolerance
END_VAR
VAR_OUTPUT
    fDpMeanKpa    : REAL;                           // 压差滑动均值 [kPa] / DP window mean [kPa]
    fTrendKpaDay  : REAL;                           // 趋势斜率 [kPa/天] / Trend slope [kPa/day]
    bClogWarn     : BOOL;                           // 堵塞预警标志（带迟滞）/ Clog warning flag
    bTrendValid   : BOOL;                           // 趋势结论有效 / Trend conclusion valid
    abMask        : BOOL;                           // 本拍压差无效掩码 / Invalid mask this scan
    bError        : BOOL;                           // 故障标志，与故障级码配对 / Fault flag
    uErrorId      : UDINT;                          // 事件码，0 = 无事件 / Event code
    eStateOut     : E_DL_ExtPhase;                  // 状态机当前态，段尾单点映射 / Phase mapped at tail
END_VAR
VAR
    _eState       : E_DL_ExtPhase := E_DL_ExtPhase.eIdle;  // 内部状态 / Internal state
    fbStatNow     : FB_DL_SignalStatistics;         // 当前窗统计实例（无条件调用）/ Current window statistics
    fbStatOld     : FB_DL_SignalStatistics;         // 快照窗统计实例（无条件调用）/ Snapshot statistics
    rtrReset      : R_TRIG;                         // 复位沿 / Reset edge
    bCfgOk        : BOOL;                           // 组态合法标志 / Configuration valid
    bDpOk         : BOOL;                           // 压差本拍有效 / DP valid this scan
    bFrozen       : BOOL;                           // 冻结合成（无效/停机）/ Frozen aggregate
    bPeriodEdge   : BOOL;                           // 周期末沿 / Period end edge
    fAccumSec     : REAL;                           // 周期累计秒 [s] / Period accumulated seconds
    fMeanNowKpa   : REAL;                           // 当前窗均值 [kPa] / Current mean [kPa]
    fMeanOldKpa   : REAL;                           // 上一周期均值快照 [kPa] / Snapshot mean [kPa]
    bWarnUp       : BOOL;                           // 预警迟滞状态（持有）/ Warning hysteresis state
    uTripCnt      : UINT;                           // 严重堵塞确认计数 [拍] / Severe confirm counter
    uFault        : UDINT;                          // 锁存故障码 / Latched fault code
    uInfo         : UDINT;                          // 信息级码 / Information code
END_VAR
VAR CONSTANT
    DL_EXT_INFMAX : REAL := 1.0E30;                 // 压差有限值幅值上限 [kPa] / DP finite bound [kPa]
    DL_EXT_MINWIN : INT := 8;                       // 趋势窗最小样本数 [样本] / Minimum window samples
END_VAR

(* === 段 0 · 实例刷新 === *)
rtrReset(CLK := bReset);                          // 每拍刷新复位沿

(* === 段 1 · 组态闸 === *)
bCfgOk := (UINT_TO_REAL(uPeriodMin) > fEps)       // 周期正域
          AND (fWarnKpa > fEps) AND (fTripKpa > fWarnKpa + fHystKpa)  // 门限不倒置且迟滞带不相交
          AND (fHystKpa > fEps) AND (fTaskCycle > fEps)
          AND (fWarnKpa = fWarnKpa) AND (fTripKpa = fTripKpa);  // NaN 自反
IF NOT bCfgOk THEN
    uFault := 16#0002_0308;                       // 故障级：组态非法
END_IF
IF rtrReset.Q AND bCfgOk THEN
    uFault := 16#0000;                            // 复位沿清锁存（解除路径可达）
    bWarnUp := FALSE;                             // 预警迟滞复位
    uTripCnt := UINT#0;                           // 严重确认计数复位
    fAccumSec := 0.0;                             // 周期累计清零
END_IF
uInfo := 16#0000;                                 // 信息码每拍清零
bDpOk := (fDpKpa = fDpKpa) AND (fDpKpa >= 0.0) AND (fDpKpa < DL_EXT_INFMAX);  // 压差 NaN 自反 + 非负域闸
abMask := NOT bDpOk;                              // 无效掩码输出
bFrozen := (NOT bDpOk) OR (NOT bFanRunning);      // 停机/无效冻结（禁把停机零流量当堵塞）
IF bFrozen AND bEnable THEN
    uInfo := 16#0002_0328;                        // 信息级：无效剔除或停机趋势冻结
END_IF

(* === 段 2 · 周期累计（先于统计实例，保快照沿同拍一致）=== *)
bPeriodEdge := FALSE;                             // 周期沿本拍重算
IF (NOT bFrozen) AND bEnable AND (uFault = 16#0000) THEN
    fAccumSec := fAccumSec + fTaskCycle;          // 非冻结拍累计
    IF fAccumSec >= UINT_TO_REAL(uPeriodMin) * 60.0 THEN
        bPeriodEdge := TRUE;                      // 周期末沿
        fAccumSec := 0.0;                         // 累计清零开新周期
    END_IF
END_IF

(* === 段 3 · 统计实例（无条件调用）与趋势折算 === *)
fbStatNow(fIn := fDpKpa,                          // 当前窗统计
          bSample := bDpOk AND bFanRunning AND (NOT bFrozen),   // 冻结拍不采（停机零流量不进窗）
          nWindow := 32,                          // 统计窗 32 样本
          bClear := rtrReset.Q);                  // 复位沿清窗
fbStatOld(fIn := fMeanNowKpa,                     // 快照窗统计（输入为均值快照）
          bSample := bPeriodEdge,                 // 周期末沿采快照
          nWindow := 8,                           // 快照窗 8 周期
          bClear := rtrReset.Q);
IF bPeriodEdge THEN
    fMeanOldKpa := fMeanNowKpa;                   // 周期末均值快照
END_IF
fDpMeanKpa := 0.0;                                // 均值缺省 0
fTrendKpaDay := 0.0;                              // 趋势缺省 0
bTrendValid := FALSE;                             // 结论缺省无效
IF fbStatNow.bStatValid AND (fbStatNow.nCount >= DL_EXT_MINWIN) THEN
    fDpMeanKpa := fbStatNow.fMean;                // 当前窗均值
    IF fbStatOld.bValid AND (fbStatOld.nCount >= 2) THEN
        fTrendKpaDay := (fDpMeanKpa - fMeanOldKpa) / (UINT_TO_REAL(uPeriodMin) / 1440.0);   // 斜率 kPa/天（分母常量防零）
        bTrendValid := TRUE;                      // 趋势结论有效
    END_IF
ELSE
    uInfo := 16#0002_0328;                        // 信息级：样本不足不出结论
END_IF

(* === 段 4 · 分级预警（预警带迟滞 / 严重持续确认升级）=== *)
IF fDpMeanKpa >= fWarnKpa THEN
    bWarnUp := TRUE;                              // 越预警门限置迟滞状态
ELSIF fDpMeanKpa < fWarnKpa - fHystKpa THEN
    bWarnUp := FALSE;                             // 回差带内解除（路径可达）
END_IF
bClogWarn := bWarnUp;                             // 预警出口
IF bDpOk AND (fDpKpa >= fTripKpa) THEN
    uTripCnt := uTripCnt + UINT#1;                // 严重堵塞确认计数
    IF uTripCnt >= uTripConfirm THEN
        uFault := 16#0002_0318;                   // 故障级：严重堵塞（锁存）
    END_IF
ELSE
    uTripCnt := UINT#0;                           // 未超严重门限计数归零
END_IF

(* === 段 5 · 主状态机（ENUM + CASE，含 ELSE 兜底）=== *)
CASE _eState OF
E_DL_ExtPhase.eIdle :
    IF uFault <> 16#0000 THEN
        _eState := E_DL_ExtPhase.eFault;          // 故障优先
    ELSIF bEnable AND bCfgOk THEN
        _eState := E_DL_ExtPhase.eWatch;          // 进监视相
    END_IF

E_DL_ExtPhase.eWatch :
    IF (uFault <> 16#0000) OR (NOT bEnable) THEN
        _eState := E_DL_ExtPhase.eFault;          // 故障/失能转出
    END_IF

E_DL_ExtPhase.eFault :
    IF uFault = 16#0000 THEN
        _eState := E_DL_ExtPhase.eIdle;           // 解锁回空闲
    END_IF

ELSE
    _eState := E_DL_ExtPhase.eFault;              // 非法状态拦截
    uFault := 16#0002_0308;                       // 故障级：相 ID 越界复用组态码段
END_CASE

(* === 段 6 · 输出映射 === *)
bError := (uFault <> 16#0000);                    // 故障标志仅由故障级码置位（R45 配对）
IF bError THEN
    uErrorId := uFault;                           // 故障级优先上报
ELSE
    uErrorId := uInfo;                            // 否则上报信息级码
END_IF
eStateOut := _eState;                             // 输出枚举段尾单点映射（N2 规则）
END_FUNCTION_BLOCK

(* ---- FB_DL_FanArrayStageCtrl.st ---- *)
(*==============================================================================
 * 组件名称 (Component)  : FB_DL_FanArrayStageCtrl
 * 所属子库 (Sublibrary) : DL_Device
 * 当前版本 (Version)    : 1.0.0
 * 兼容性 (Platform)     : CODESYS 3.5 / TwinCAT 3 / 汇川 InoProShop / Machine Expert
 *                         仅依赖纯 IEC 61131-3 标准元素，零厂商方言
 * 功能描述 (Function)   : N+1 风机阵列分级启停：按需求级数对称加/减机，
 *                         每 tick 至多切换 1 台（加机选运行小时最少者、减机选
 *                         运行小时最多者，轮值均衡）；tMinRun/tMinStop 闸门
 *                         防频繁启停；需求级数钳位 [0, 台数-1] 预留 1 台备机。
 * 溯源 (Origin)         : 道莅 clean-room 防御性实现
 * 本文件内含 (Contains) : TYPE E_DL_FanArrErr / FUNCTION_BLOCK FB_DL_FanArrayStageCtrl
 * 依赖 (Depends)        : 无 DL_ 内部依赖；Standard.library TON 实例
 * 红线自检 (Redline)    : 无外部全局变量、无硬件地址直引 ｜ 全变量中英双语同行注释
 *                         数组下界常量提取 + 防越界 ｜ 枚举成员全部显式赋值
 *                         TON 实例每周期无条件调用（仅 IN 条件化）｜ CASE 含 ELSE 兜底
 * 错误码表 (Codes)      : 16#0003_038E 就绪
 *                         16#0003_038F 信息级 台数越界(已钳制 8)
 *                         16#0003_0390 信息级 需求级数越界(已钳制)
 *                         16#0003_0391 信息级 最短时序未满足(等待中)
 *                         16#0003_0392 信息级 运行小时数据全零(轮值退化按顺序)
 * 修订历史 (Revision)   : 2026-11-17  v1.0.0  首版入库 · R27 · 阶段三批 2
 * 验收向量 (Acceptance) : total=4, req=3, 全部停机 → 逐拍加机至 3 台；
 *                         req=4 → 钳 3（预留备机）0390；切换后 tMinRun 内再要求切换 → 0391
 *============================================================================*)

(*-----------------------------------------------------------------------------
 * 枚举: E_DL_FanArrErr（归属 DL_Device，与 FB_DL_FanArrayStageCtrl 同文件）
 *----------------------------------------------------------------------------*)
TYPE E_DL_FanArrErr :
(
    eReady       := 16#0003_038E,   // 就绪 / Ready
    eTotalClamp  := 16#0003_038F,   // 信息级：台数越界已钳制 / Info: total clamped
    eStageClamp  := 16#0003_0390,   // 信息级：需求级数越界已钳制 / Info: stage request clamped
    eGateWait    := 16#0003_0391,   // 信息级：最短时序未满足（等待）/ Info: min-run gate waiting
    eHrsAllZero  := 16#0003_0392    // 信息级：运行小时全零，轮值退化按顺序 / Info: all run-hours zero, round-robin degenerated
);
END_TYPE

(*==============================================================================
 * 功能块: FB_DL_FanArrayStageCtrl
 * 调用约定: 每个扫描周期无条件调用一次；aNRunHrs 由调用方按索引注入。
 *============================================================================*)
FUNCTION_BLOCK FB_DL_FanArrayStageCtrl
VAR_INPUT
    aNRunHrs     : ARRAY[1..8] OF UDINT;   // 各风机累计运行小时 [小时] / Run hours per fan [h]
    uStageReq    : UINT;                   // 需求级数 [台]，有效域 0~8 / Requested stage count [fans]
    uFanTotal    : UINT;                   // 装机台数 [台]，有效域 1~8 / Installed fan count [fans]
    tMinRun      : TIME := T#60S;          // 最短运行时长 [秒] / Minimum run time [s]
    tMinStop     : TIME := T#60S;          // 最短停机时长 [秒] / Minimum stop time [s]
END_VAR
VAR_OUTPUT
    auFanCmd     : ARRAY[1..8] OF BOOL;    // 各风机启停指令 / Fan start/stop commands
    uStageAct    : UINT;                   // 实际运行级数 [台] / Actual running stage count [fans]
    eErr         : E_DL_FanArrErr;         // 错误码 / Error code
END_VAR
VAR
    tonGateRun   : TON;                    // 最短运行闸门定时器（无条件调用）/ Min-run gate timer
    tonGateStop  : TON;                    // 最短停机闸门定时器（无条件调用）/ Min-stop gate timer
    bGateArmed   : BOOL;                   // 闸门武装标志（切换后置位）/ Gate armed flag, set on any switch
    bSwitchCycle : BOOL;                   // 本拍为切换拍（定时器 IN 强制断开以复位）/ TRUE on the switch scan, forces timer reset
    uTotalUse    : UINT;                   // 生效台数（钳位后）[台] / Effective installed count [fans]
    uStageUse    : UINT;                   // 生效需求级数（钳位后）[台] / Effective requested stage [fans]
    uIdxBest     : UINT;                   // 候选切换风机索引 [台序] / Candidate fan index for switching
    uHoursZero   : INT;                    // 运行小时为零的风机计数 [台] / Count of fans with zero hours
    i            : INT;                    // 数组循环索引 / Array loop index
    nPickHrs     : UDINT;                  // 候选比较基准小时 [小时] / Candidate comparison hours baseline [h]
    bInit        : BOOL;                   // 首扫初始化标志 / First-scan init flag
END_VAR
VAR CONSTANT
    DL_FAN_IDX_MAX   : INT  := 8;          // 阵列容量上限（数组下界常量提取）/ Array capacity upper bound
    DL_FAN_TOTAL_MAX : UINT := 8;          // 装机台数上限 [台] / Installed count upper bound [fans]
    DL_FAN_RESERVE   : UINT := 1;          // N+1 预留备机数 [台] / Reserved standby count [fans]
    DL_FAN_CNT_SAT   : UINT := 65535;      // 级数输出饱和值 [台] / Stage output saturation [fans]
END_VAR

(*------------------------------------------------------------------------------
 * 段 1｜TON 实例每周期无条件调用（仅 IN 条件化）：切换拍强制断流以复位计时
 *----------------------------------------------------------------------------*)
tonGateRun(IN := bGateArmed AND NOT bSwitchCycle, PT := tMinRun);    // 运行闸计时 / min-run gate timing
tonGateStop(IN := bGateArmed AND NOT bSwitchCycle, PT := tMinStop);  // 停机闸计时 / min-stop gate timing

(*------------------------------------------------------------------------------
 * 段 2｜首扫初始化：按当前台数同步指令数组（默认全停）
 *----------------------------------------------------------------------------*)
IF NOT bInit THEN
    FOR i := 1 TO DL_FAN_IDX_MAX DO
        auFanCmd[i] := FALSE;                        // 默认全停 / default all stopped
    END_FOR
    bInit := TRUE;                                   // 首扫完成 / first scan done
END_IF

(*------------------------------------------------------------------------------
 * 段 3｜台数钳位（信息级）：装机台数钳 [1, 8]
 *----------------------------------------------------------------------------*)
eErr := E_DL_FanArrErr.eReady;                       // 预置就绪 / preset ready
uTotalUse := uFanTotal;                              // 台数工作副本 / total working copy
IF uTotalUse > DL_FAN_TOTAL_MAX THEN
    uTotalUse := DL_FAN_TOTAL_MAX;                   // 台数上限钳位 / total capped
    eErr := E_DL_FanArrErr.eTotalClamp;              // 信息级：台数越界 / info: total clamped
ELSIF uTotalUse < 1 THEN
    uTotalUse := 1;                                  // 台数下限钳位 / total floored
    eErr := E_DL_FanArrErr.eTotalClamp;              // 信息级：台数越界 / info: total clamped
END_IF

(*------------------------------------------------------------------------------
 * 段 4｜需求级数钳位 [0, 台数-1]（预留 1 台备机，N+1 纪律）
 *----------------------------------------------------------------------------*)
uStageUse := uStageReq;                              // 需求工作副本 / request working copy
IF uStageUse > (uTotalUse - DL_FAN_RESERVE) THEN
    uStageUse := uTotalUse - DL_FAN_RESERVE;         // 级数上限钳位（预留备机）/ stage capped, standby reserved
    IF eErr = E_DL_FanArrErr.eReady THEN
        eErr := E_DL_FanArrErr.eStageClamp;          // 信息级：需求级数越界 / info: stage clamped
    END_IF
END_IF

(*------------------------------------------------------------------------------
 * 段 5｜轮值数据体检：运行小时全零计数（全零则轮值退化按索引顺序）
 *----------------------------------------------------------------------------*)
uHoursZero := 0;                                     // 全零计数清零 / zero-hours count reset
FOR i := 1 TO UINT_TO_INT(uTotalUse) DO
    IF aNRunHrs[i] = 0 THEN
        uHoursZero := uHoursZero + 1;                // 全零风机计数 [台] / count zero-hour fans
    END_IF
END_FOR
IF uHoursZero = UINT_TO_INT(uTotalUse) THEN
    IF eErr = E_DL_FanArrErr.eReady THEN
        eErr := E_DL_FanArrErr.eHrsAllZero;          // 信息级：轮值退化按顺序 / info: round-robin degenerated
    END_IF
END_IF

(*------------------------------------------------------------------------------
 * 段 6｜每 tick 至多切换 1 台：加机选运行小时最少者，减机选运行小时最多者
 *----------------------------------------------------------------------------*)
uIdxBest := 0;                                       // 候选索引清零（0 = 无候选）/ candidate reset, 0 means none
nPickHrs := 0;                                       // 候选基准清零 / baseline reset
IF uStageAct > uStageUse THEN
    // 减机：在运行台中选运行小时最多者（轮值均衡）/ shed: pick running fan with most hours
    IF bGateArmed AND NOT tonGateRun.Q THEN
        IF eErr = E_DL_FanArrErr.eReady THEN
            eErr := E_DL_FanArrErr.eGateWait;        // 信息级：最短时序未满足 / info: gate waiting
        END_IF
    ELSE
        nPickHrs := 0;                               // 最多小时基准从 0 起比 / start from zero for max search
        FOR i := 1 TO UINT_TO_INT(uTotalUse) DO
            IF auFanCmd[i] THEN
                IF (uIdxBest = 0) OR (aNRunHrs[i] >= nPickHrs) THEN
                    uIdxBest := INT_TO_UINT(i);      // 候选更新（运行最久者）/ candidate updated, most-run fan
                    nPickHrs := aNRunHrs[i];         // 基准更新 / baseline updated
                END_IF
            END_IF
        END_FOR
    END_IF
ELSIF uStageAct < uStageUse THEN
    // 加机：在停机台中选运行小时最少者（轮值均衡）/ add: pick stopped fan with least hours
    IF bGateArmed AND NOT tonGateStop.Q THEN
        IF eErr = E_DL_FanArrErr.eReady THEN
            eErr := E_DL_FanArrErr.eGateWait;        // 信息级：最短时序未满足 / info: gate waiting
        END_IF
    ELSE
        nPickHrs := 16#FFFF_FFFF;                    // 最少小时基准从满值起比 / start from max for min search
        FOR i := 1 TO UINT_TO_INT(uTotalUse) DO
            IF NOT auFanCmd[i] THEN
                IF aNRunHrs[i] <= nPickHrs THEN
                    uIdxBest := INT_TO_UINT(i);      // 候选更新（停机最久者近似为小时最少）/ candidate updated, least-run fan
                    nPickHrs := aNRunHrs[i];         // 基准更新 / baseline updated
                END_IF
            END_IF
        END_FOR
    END_IF
END_IF

(*------------------------------------------------------------------------------
 * 段 7｜执行切换：切换拍置武装标志并强制定时器断流复位
 *----------------------------------------------------------------------------*)
bSwitchCycle := FALSE;                               // 切换拍标志默认 FALSE / switch-scan flag defaults FALSE
IF uIdxBest > 0 THEN
    auFanCmd[UINT_TO_INT(uIdxBest)] := NOT auFanCmd[UINT_TO_INT(uIdxBest)];   // 执行切换 / execute the switch
    bGateArmed := TRUE;                              // 闸门武装 / gate armed
    bSwitchCycle := TRUE;                            // 切换拍标志（下拍定时器重新计时）/ switch scan flag
END_IF

(*------------------------------------------------------------------------------
 * 段 8｜实际级数统计与数组上界外指令清扫（防越界残留）
 *----------------------------------------------------------------------------*)
uStageAct := 0;                                      // 实际级数清零 / actual stage reset
FOR i := 1 TO DL_FAN_IDX_MAX DO
    IF i > UINT_TO_INT(uTotalUse) THEN
        auFanCmd[i] := FALSE;                        // 容量外指令强制撤销（防越界残留）/ force FALSE beyond capacity
    ELSIF auFanCmd[i] THEN
        uStageAct := uStageAct + 1;                  // 运行台数累加 [台] / count running fans
    END_IF
END_FOR
IF uStageAct > DL_FAN_CNT_SAT THEN
    uStageAct := DL_FAN_CNT_SAT;                     // 级数饱和防护 / stage saturation guard
END_IF
END_FUNCTION_BLOCK

(* ---- FB_DL_FanBeltSlipDetect.st ---- *)
(*
  Component : FB_DL_FanBeltSlipDetect
  Category  : DL_Device
  Type      : FB
  Version   : 1.0.0
  CodeSeg   : 16#03_1_01
  Summary   : 风机皮带打滑判据：转速比（风扇/电机）偏差速率越阈判打滑，锁存告警并带维护提醒计数。
              Fan belt slip detection: speed-ratio deviation rate over threshold latches the alarm with a maintenance counter.
  溯源声明  : 道莅自研 clean-room
  边界安全  : 电机转速正域闸（> eps 防比值除零）；输入非有限（NaN 自反 + Inf 上限）拦截；
              采样窗时长域闸（tWinMs > 0，防 dt 为零除零）；比值偏差速率比较带容差；
              TON 实例每拍无条件刷新且自复位振荡（IN := NOT ton.Q）；锁存有可达恢复清码路径。
  复用      : 无
*)

FUNCTION_BLOCK FB_DL_FanBeltSlipDetect
VAR_INPUT
    bRun       : BOOL;                  (* 监视使能 · Enable *)
    fMotRpm    : LREAL;                 (* 电机转速 [rpm] · Motor speed *)
    fFanRpm    : LREAL;                 (* 风扇转速 [rpm] · Fan speed *)
    fRatioNom  : LREAL := 1.0;          (* 额定风扇/电机转速比 [比值] · Nominal speed ratio *)
    fDevRateTh : LREAL := 0.02;         (* 打滑判据：比值偏差速率阈 [比值/s] · Slip rate threshold *)
    tWinMs     : TIME  := T#1000MS;     (* 采样窗时长 [ms]，禁魔法数 · Sample window *)
    tClearMs   : TIME  := T#5000MS;     (* 恢复清码持续时长 [ms] · Recovery clear duration *)
    fEps       : LREAL := 1.0E-6;       (* 浮点判零容差 [实数域] · Floating zero tolerance *)
END_VAR
VAR_OUTPUT
    bSlip      : BOOL;                  (* 打滑锁存告警 · Latched slip alarm *)
    fRatioNow  : LREAL;                 (* 当前转速比 [比值] · Current speed ratio *)
    fDevRate   : LREAL;                 (* 比值偏差速率 [比值/s] · Ratio deviation rate *)
    nSlipCount : UDINT;                 (* 打滑事件累计 [次]，防回卷 · Slip event count *)
    bMaintHint : BOOL;                  (* 维护提醒（累计超阈）· Maintenance hint *)
    bError     : BOOL;                  (* 故障标志，与故障码配对 · Fault flag paired with codes *)
    uErrorId   : UDINT;                 (* 事件码 16#0000_0101，0 无事件 · Event code *)
END_VAR
VAR
    uCode    : WORD;    (* 码位暂存，每拍重算 [码] · Code staging *)
    tonWin   : TON;     (* 采样窗节拍定时器 [ms]，自复位振荡 · Sample window timer, self-reset *)
    tonClr   : TON;     (* 恢复清码定时器 [ms] · Recovery clear timer *)
    bSigOk   : BOOL;    (* 输入有效标志 · Input validity flag *)
    bTick    : BOOL;    (* 采样窗到点脉冲 [脉冲] · Sample tick pulse *)
    fDtS     : LREAL;   (* 采样窗秒值 [s]，一次导出 · Window seconds derived once *)
    fRatioPrv: LREAL;   (* 上窗比值快照 [比值] · Previous ratio snapshot *)
    bSlipPrv : BOOL;    (* 上拍锁存快照，事件沿判据 · Previous latch snapshot *)
    nSlipCnt2: INT;     (* 连续越阈窗数 [窗] · Consecutive over-threshold windows *)
    nCycles  : UDINT;   (* 有效采样窗计数 [窗]，防回卷 · Sampled window count *)
END_VAR
VAR CONSTANT
    DL_FBS_WRAP  : UDINT := 4294967290; (* 计数防回卷余量 [次] · Counter wrap guard *)
    DL_FBS_HINTN : UDINT := 3;          (* 维护提醒事件阈 [次] · Maintenance hint threshold *)
END_VAR

(* === 段 0 · 实例刷新（每拍无条件，红线 7）=== *)
tonWin(IN := NOT tonWin.Q, PT := tWinMs);       // 采样窗自复位振荡 / Self-reset oscillating window
tonClr(IN := bSigOk AND (NOT bSlip) AND (nSlipCnt2 = 0), PT := tClearMs);
                                                // 恢复计时：比值正常且无越阈时计时 / Recovery timing
bTick := tonWin.Q;                              // 窗到点脉冲 / Tick pulse

(* === 段 1 · 输入校验与量程闸 === *)
uCode := 16#0000;                       // 每拍清码（可达清零基线）/ Clear codes each scan
bSigOk := (fMotRpm = fMotRpm) AND (fFanRpm = fFanRpm) AND (fRatioNom = fRatioNom)
          AND (ABS(fMotRpm) < 1.0E308) AND (ABS(fFanRpm) < 1.0E308)     // 非有限拦截 / Non-finite guard
          AND (fMotRpm > fEps) AND (fRatioNom > fEps)                   // 转速/比值正域闸 / Positive domain
          AND (tWinMs > T#0MS);                                         // 窗时长正域闸 / Window duration gate
IF fDtS < fEps THEN
    fDtS := DINT_TO_LREAL(TIME_TO_DINT(tWinMs)) / 1000.0;   // 窗秒值一次导出 / Derive window seconds once
END_IF
IF NOT bSigOk THEN
    uCode := 16#0101;                   // 故障级：输入域外，判据冻结 / Fault: input domain invalid
END_IF

(* === 段 2 · 主逻辑：比值-偏差速率判据 === *)
IF bSigOk THEN
    fRatioNow := fFanRpm / fMotRpm;     // 当前转速比（分母已闸）/ Current ratio
    IF bTick THEN
        fDevRate := (fRatioNow - fRatioPrv) / fDtS;     // 偏差速率 [比值/s]，先算后存快照 / Rate first, then snapshot
        fRatioPrv := fRatioNow;         // 快照更新 / Update the snapshot
        IF ABS(fDevRate) > fDevRateTh THEN
            nSlipCnt2 := nSlipCnt2 + 1; // 连续越阈窗数累加 / Count over-threshold windows
        ELSE
            nSlipCnt2 := 0;             // 正常窗清计数 / Clear on a normal window
        END_IF
        IF nCycles < DL_FBS_WRAP THEN
            nCycles := nCycles + 1;     // 有效窗计数 / Count valid windows
        END_IF
    END_IF
    IF nSlipCnt2 >= 2 THEN              // 连续 2 窗越阈才判打滑（防单拍毛刺）/ Two windows to latch
        bSlip := TRUE;                  // 打滑锁存 / Latch the slip
    END_IF
    IF tonClr.Q THEN                    // 恢复条件持续满足 → 可达清锁存 / Reachable clear path
        bSlip := FALSE;                 // 解除锁存 / Release the latch
        fDevRate := 0.0;                // 速率复位 / Reset the rate
    END_IF
END_IF

(* === 段 3 · 输出映射与故障码 === *)
IF bSlip AND (NOT bSlipPrv) THEN
    IF nSlipCount < DL_FBS_WRAP THEN
        nSlipCount := nSlipCount + 1;   // 打滑事件沿计数 / Count slip events on the edge
    END_IF
END_IF
bSlipPrv := bSlip;                      // 锁存快照 / Latch snapshot
bMaintHint := (nSlipCount >= DL_FBS_HINTN);     // 维护提醒 / Maintenance hint
bError := bSlip OR (uCode <> 16#0000);  // 故障标志：打滑或域外 / Fault flag
IF bSlip THEN
    uErrorId := WORD_TO_UDINT(16#0101); // 码位 16#0000_0101 打滑锁存 / Slip latch code
ELSE
    uErrorId := WORD_TO_UDINT(uCode);   // 域外码或零 / Domain code or zero
END_IF
END_FUNCTION_BLOCK

(* ---- FB_DL_FanBeltSlipDiag.st ---- *)
(*==============================================================================
 * 组件名称 (Component)  : FB_DL_FanBeltSlipDiag
 * 溯源说明 (Provenance) : 道莅 clean-room 防御性实现（Building 泵风机族深化）
 * 所属子库 (Sublibrary) : DL_Device / FanDiag
 * 当前版本 (Version)    : 1.0.0
 * 兼容性   (Platform)   : CODESYS 3.5 / TwinCAT 3 / 汇川 InoProShop；
 *                         纯 IEC 61131-3（第 3 版），仅用标准库 TON
 * 组件分类 (Category)   : 功能块（FUNCTION_BLOCK）· 风机皮带打滑诊断
 * 功能一句话 (Summary)  : 电机/叶轮转速比监视 + 确认延时 + 叶轮停转判据。
 * 边界与安全 (Boundary) : ①电机转速小于 1 rpm 不判定（防除零，规格口径）；
 *                         ②bMotorRun=FALSE 清确认（停机撤销判定）；
 *                         ③叶轮近零而电机运行 → 叶轮停转码；
 *                         ④转速负值或非有限 → 输入非法码；
 *                         ⑤确认 TON 无条件周期刷新；
 *                         ⑥转速比按 1:1 皮带传动基准（倍率差异属调用方换算）。
 * 错误码    : 16#0003_0381 转速比超差确认（打滑）——故障级（持续态）
 *             16#0003_0382 叶轮停转而电机运行——故障级（持续态）
 *             16#0003_0383 输入非法（负转速或非有限）——故障级（持续态）
 * 码位总账  : 16#0003_0381 用 / 16#0003_0382 用 / 16#0003_0383 用
 * 修改记录  : v1.0.0 R26 初版
 *==============================================================================*)
FUNCTION_BLOCK FB_DL_FanBeltSlipDiag
VAR_INPUT
    fMotorRpm : LREAL; // 电机转速 [rpm] / Motor speed [rpm]
    fFanRpm   : LREAL; // 叶轮转速 [rpm] / Fan wheel speed [rpm]
    fRatioTol : LREAL; // 转速比容差 [%] / Speed ratio tolerance [%]
    tConfirm  : TIME;  // 打滑确认延时 [ms] / Slip confirm delay [ms]
    bMotorRun : BOOL;  // 电机运行反馈 / Motor running feedback
END_VAR
VAR_OUTPUT
    bSlip        : BOOL; // 打滑特征成立（计时中）/ Slip signature active
    bSlipConfirm : BOOL; // 打滑确认（延时满足）/ Slip confirmed
    fRatio       : LREAL; // 电机/叶轮转速比 / Motor-to-fan speed ratio
    eErr         : UDINT; // 本周期错误码，0=无错 / Error code this cycle, 0 = none
END_VAR
VAR CONSTANT
    cMinRpm : LREAL := 1.0; // 判定最小电机转速 [rpm] / Minimum judgeable motor speed
END_VAR
VAR
    tonSlip : TON;   // 打滑确认定时器（无条件刷新）/ Slip confirm timer
    bInSlip : BOOL;  // 打滑域内判据 / In-slip-domain predicate
    bInOk   : BOOL;  // 输入合法性 / Input legality
    fMotGrd : LREAL; // 电机转速守卫副本 / Motor speed guard copy
    fFanGrd : LREAL; // 叶轮转速守卫副本 / Fan speed guard copy
    fSlip   : LREAL; // 比值偏离量 [%] / Ratio deviation [%]
END_VAR

// ---------- 实时守卫副本 ----------
fMotGrd := fMotorRpm;
fFanGrd := fFanRpm;

// ---------- 输入合法性：负转速或非有限拒判 ----------
bInOk := bMotorRun AND (fMotGrd >= 0.0) AND (fFanGrd >= 0.0)
     AND (fMotGrd = fMotGrd) AND (fFanGrd = fFanGrd);
IF NOT bInOk THEN
    IF bMotorRun AND ((fMotGrd < 0.0) OR (fFanGrd < 0.0)
       OR (fMotGrd <> fMotGrd) OR (fFanGrd <> fFanGrd)) THEN
        eErr := 16#0003_0383;                 // 输入非法码 / Illegal input code
    ELSE
        eErr := 0;                            // 停机不置码（正常撤销）/ Stopped, no code
    END_IF
END_IF

// ---------- 转速比计算：电机转速小于 1 rpm 不判定（防除零） ----------
IF bInOk AND (fMotGrd >= cMinRpm) THEN
    IF fFanGrd > 0.0 THEN
        fRatio := fMotGrd / fFanGrd;          // 除法前判零 / Zero-guarded divide
        fSlip := (fRatio - 1.0) * 100.0;      // 偏离百分比 / Deviation percent
        IF fSlip < 0.0 THEN
            fSlip := -fSlip;                  // 绝对偏离 / Absolute deviation
        END_IF
        bInSlip := fSlip > fRatioTol;         // 超差判据 / Over-tolerance predicate
    ELSE
        fRatio := 0.0;                        // 叶轮停转比值缺省 / Stalled wheel default
        bInSlip := FALSE;
        eErr := 16#0003_0382;                 // 叶轮停转码 / Wheel stall code
    END_IF
ELSE
    fRatio := 0.0;                            // 不判定缺省 / Not-judged default
    bInSlip := FALSE;
END_IF

// ---------- 无条件周期刷新：打滑确认定时器 ----------
tonSlip(IN := bInSlip, PT := tConfirm);
bSlip := tonSlip.IN;                          // 计时中特征 / Signature while timing
IF tonSlip.Q THEN
    bSlipConfirm := TRUE;                     // 确认成立 / Confirmed
    eErr := 16#0003_0381;                     // 超差确认码 / Over-tolerance confirm code
ELSE
    bSlipConfirm := FALSE;                    // 未确认即撤销 / Withdrawn if unconfirmed
END_IF

END_FUNCTION_BLOCK

(* ---- FB_DL_FanVfdBypassSwap.st ---- *)
(*
  ==================================================================
  组件名 Component  : FB_DL_FanVfdBypassSwap
  分类   Category   : DL_Device
  复杂度 Complexity  : cx4
  版本   Version    : 1.0.0
  功能   Purpose    : 单台风机变频 → 工频旁通切换顺控。相位机 eIdle → eStopVfd →
                      eWaitSpinDown → eCloseBypass → eRunDurance → eStable / eFault；
                      任何中间态严格双断（bVfdRun 与 bBypassRun 不同拍同为真）；
                      含降速阈值判据、切换最小间隔窗 tGapMin、旁通接触器确认反馈
                      bBypassFb、失败重试 nRetryMax 与超时 eSwapTimeout。
  来源   Source     : t2-2-lbp
  溯源   Origin     : IEC 61131-3 标准语义的道莅防御性实现；变频 / 工频旁通切换
                      时序为通用电气传动语义，clean-room 自研实现，未复制任何
                      闭源代码行。
  平台   Platform   : 纯 IEC 61131-3（TON / R_TRIG / LREAL，无私有库）
  作者   Author     : 道莅代码库 · PLC 编程专家（R56）
  ------------------------------------------------------------------
  同拍多窗配比约束（R100）：五个窗职责分离 —— tStopTo 判变频反馈消失（短），
                      tGapMin 切换最小间隔（中），tSpinMax 降速总窗（长），
                      tCloseTo 旁通反馈确认窗，tStableMin 稳定驻留窗；
                      配比约束 tSpinMax > tGapMin 在组态域闸内直接判故障，
                      其余各窗互斥（每窗 IN 串本相闸），任一时刻只有一个窗在计时。
  边界 Boundary     :
                      一 本件只出切换命令与诊断，不做接触器本体驱动、不写变频器参数
                         （属主边界）；
                      二 互斥不变量：bVfdRun 与 bBypassRun 恒不同拍为真（结构性成立，
                         出口为相位派生电平）；
                      三 相级看门狗使能只用「相驻留」本身（R145），不叠加业务条件补集；
                      四 故障锁存解除路径 = bReset 上升沿（唯一路径，头注释声明，R188）；
                      五 eWaitSpinDown 相退出条件 ≥2 条（转速达标 / 超时 / 失能，R98）；
                      六 无全局变量、无外部变量声明、无物理地址寻址。
  输出契约 Output contract:
                      bVfdRun / bBypassRun 为相位派生命令电平，相外恒假；
                      bBothOff 为双断指示（两命令均假的派生量）；
                      eFault 为锁存回放；ePhaseBad 为非法相位兜底专用成员（R128）。
  修订记录 Revision  :
    2026-11-20  v1.0.0  R56 首版（批 3 · 序号 12）
  ==================================================================
*)

TYPE E_DL_FbsPhase :
(
    eIdle        := 0,  // 空闲：变频运行保持，等切换申请 / idle, the VFD holds and waits for a swap request
    eStopVfd     := 10, // 停变频：撤变频命令等反馈消失 / stopping, the VFD command is withdrawn and the feedback awaited
    eWaitSpinDown:= 20,  // 等降速：转速阈值 + 最小间隔窗双判 / waiting, the speed threshold and the gap window
    eCloseBypass := 30,  // 关旁通：出旁通命令等反馈确认 / closing, the bypass command waits for the feedback
    eRunDurance  := 40, // 稳定中：旁通保持，驻留稳定窗 / running in, the bypass holds through the stability window
    eStable      := 50, // 已稳定：旁通运行，监视反馈 / stable, the bypass runs with feedback watch
    eFault       := 90  // 故障：成因锁存，双断 / fault, the cause is latched with both commands off
);
END_TYPE

TYPE E_DL_FbsFault :
(
    eNone          := 0, // 无成因 / no cause
    eSwapTimeout   := 1, // 切换超时（停变频或降速窗耗尽，故障级，与 bError 配对）/ the swap timed out, fault grade paired with bError
    eFbLost        := 2, // 旁通反馈丢失（故障级，与 bError 配对）/ the bypass feedback was lost, fault grade paired with bError
    eRetryExhausted := 3, // 重试用尽（故障级，与 bError 配对）/ the retries were exhausted, fault grade paired with bError
    eCfgIllegal    := 4, // 组态非法（故障级，与 bError 配对）/ illegal configuration, fault grade paired with bError
    ePhaseBad      := 5  // 非法相位兜底（故障级，与 bError 配对）/ illegal phase fallback, fault grade paired with bError
);
END_TYPE

FUNCTION_BLOCK FB_DL_FanVfdBypassSwap
VAR_INPUT
    bEnable    : BOOL := TRUE;    // 使能，失能时停顺控回空闲 [-] / enable, the sequence stops when disabled
    bReset     : BOOL := FALSE;   // 复位上升沿清故障锁存与重试计数 [-] / reset rising edge clears the fault latch and the retry count
    bStartSwap : BOOL := FALSE;   // 切换申请脉冲，上升沿受理 [-] / the swap request pulse, accepted on the rising edge
    bAbort     : BOOL := FALSE;   // 中止（电平），任何中间态立即双断回空闲 [-] / abort level, any middle phase goes both off and back to idle
    bVfdFb     : BOOL := TRUE;    // 变频运行反馈 [-] / the VFD running feedback
    bBypassFb  : BOOL := FALSE;   // 旁通接触器确认反馈 [-] / the bypass contactor feedback
    fSpeed     : LREAL := 0.0;    // 风机实际转速 [转每分] / the actual fan speed [rpm]
    fSpeedMin  : LREAL := 50.0;   // 旁通投入转速阈值 [转每分]，域 大于零 / the bypass engagement speed threshold [rpm], domain above zero
    nRetryMax  : INT := 2;        // 旁通重试上限 [次]，域 0..9 / the retry ceiling [count], domain zero to nine
    tStopTo    : TIME := T#10S;   // 变频反馈消失窗 [毫秒]，域 大于零 / the VFD feedback drop window [millisecond], domain above zero
    tGapMin    : TIME := T#2S;    // 切换最小间隔窗 [毫秒]，域 大于零 / the minimum swap gap window [millisecond], domain above zero
    tSpinMax   : TIME := T#60S;   // 降速总窗 [毫秒]，域 大于 tGapMin / the spin down window [millisecond], above the gap
    tCloseTo   : TIME := T#5S;    // 旁通反馈确认窗 [毫秒]，域 大于零 / the bypass feedback confirm window [millisecond], domain above zero
    tStableMin : TIME := T#10S;   // 稳定驻留窗 [毫秒]，域 大于零 / the stability dwell window [millisecond], domain above zero
END_VAR
VAR_OUTPUT
    bVfdRun    : BOOL := FALSE;  // 变频运行保持命令（相位派生电平）[-] / the VFD hold command, a phase derived level
    bBypassRun : BOOL := FALSE;  // 旁通运行命令（相位派生电平）[-] / the bypass run command, a phase derived level
    bBothOff   : BOOL := TRUE;   // 双断指示（两命令均假）[-] / the both off indicator
    nRetry     : INT := 0;       // 当前重试次数 [次] / the current retry count [count]
    ePhase     : E_DL_FbsPhase := E_DL_FbsPhase.eIdle; // 相位出口 [枚举] / phase outlet [enum]
    eFault     : E_DL_FbsFault := E_DL_FbsFault.eNone; // 成因出口，锁存回放 [枚举] / cause outlet replayed from the latch [enum]
    bError     : BOOL := FALSE;  // 故障锁存标志 [-] / fault latch flag
END_VAR
VAR
    rtSwap     : R_TRIG; // 切换申请沿检测，段 0 无条件刷新 / swap request edge, refreshed unconditionally in segment zero
    rtReset    : R_TRIG; // 复位沿检测，段 0 无条件刷新 / reset edge, refreshed unconditionally in segment zero
    tonStop    : TON;    // 变频反馈消失窗，段 0 无条件刷新 / the VFD feedback drop window, refreshed unconditionally
    tonGap     : TON;    // 切换最小间隔窗，段 0 无条件刷新 / the minimum gap window, refreshed unconditionally
    tonSpin    : TON;    // 降速总窗，段 0 无条件刷新 / the spin down window, refreshed unconditionally
    tonClose   : TON;    // 旁通反馈确认窗，段 0 无条件刷新 / the feedback confirm window, refreshed unconditionally
    tonStable  : TON;    // 稳定驻留窗，段 0 无条件刷新 / the stability dwell window, refreshed unconditionally
    _ePhase    : E_DL_FbsPhase := E_DL_FbsPhase.eIdle; // 内部相位，CASE 唯一写入目标 / internal phase, the only CASE write target
    _eFaulC    : E_DL_FbsFault := E_DL_FbsFault.eNone; // 故障级成因，锁存至复位沿 / fault cause, latched until the reset edge
    _bFault    : BOOL := FALSE; // 故障锁存位 [-] / fault latch bit
    _bInit     : BOOL := FALSE; // 首扫初始化完成标志（R310）/ first scan initialisation flag
    _bCfgBad   : BOOL := FALSE; // 组态非法判定 [-] / the illegal configuration verdict
    _nRetry    : INT := 0;      // 重试计数工作值 [次] / the retry count working value [count]
    _nRetryUse : INT := 2;      // 钳定后的重试上限 [次] / the clamped retry ceiling [count]
END_VAR

// 段 0｜定时器与沿检测无条件周期刷新（禁入分支），IN 只串相位闸与故障闸（FB50-1）/ segment 0, unconditional refresh, no instance call inside a branch
rtSwap(CLK := bStartSwap); // 切换申请沿 / the swap request edge
rtReset(CLK := bReset); // 复位沿 / the reset edge
tonStop(IN := (_ePhase = E_DL_FbsPhase.eStopVfd) AND (NOT _bFault), PT := tStopTo); // 变频反馈消失窗 / the VFD feedback drop window
tonGap(IN := (_ePhase = E_DL_FbsPhase.eWaitSpinDown) AND (NOT bVfdFb) AND (NOT _bFault), PT := tGapMin); // 最小间隔窗，自变频反馈消失起计 / the gap window from the feedback drop
tonSpin(IN := (_ePhase = E_DL_FbsPhase.eWaitSpinDown) AND (NOT _bFault), PT := tSpinMax); // 降速总窗 / the spin down window
tonClose(IN := (_ePhase = E_DL_FbsPhase.eCloseBypass) AND (NOT _bFault), PT := tCloseTo); // 旁通反馈确认窗 / the feedback confirm window
tonStable(IN := (_ePhase = E_DL_FbsPhase.eRunDurance) AND (NOT _bFault), PT := tStableMin); // 稳定驻留窗 / the stability dwell window

// 段 1｜首扫初始化（R310）/ segment 1, first scan initialisation
IF NOT _bInit THEN // 首扫一拍 / the very first scan
    _bInit := TRUE; // 置首扫完成标志 / raise the first scan flag
    _ePhase := E_DL_FbsPhase.eIdle; // 相位从空闲起步 / the phase starts from idle
    _eFaulC := E_DL_FbsFault.eNone; // 故障级成因清零 / clear the fault cause
    _bFault := FALSE; // 故障锁存清零 / clear the fault latch
    _nRetry := 0; // 重试计数清零 / clear the retry count
END_IF

// 段 2｜复位沿作用域：清锁存 / 迁相位 / 清重试计数（三项逐项声明）/ segment 2, reset edge scope declared item by item
IF rtReset.Q THEN // 复位沿 / the reset edge
    _bFault := FALSE; // 作用域一：清故障锁存 / scope one, clear the fault latch
    _eFaulC := E_DL_FbsFault.eNone; // 作用域一：清故障级成因 / scope one, clear the fault cause
    _ePhase := E_DL_FbsPhase.eIdle; // 作用域二：迁回空闲相 / scope two, migrate back to idle
    _nRetry := 0; // 作用域三：清重试计数 / scope three, clear the retry count
END_IF

// 段 3｜组态域闸（R151 全覆盖，含 R100 配比约束）/ segment 3, the configuration gate with the window pairing constraint
_bCfgBad := FALSE; // 组态非法预置假 / preset the illegal configuration verdict to false
IF (fSpeedMin <= 0.0) OR (fSpeedMin <> fSpeedMin) OR ((fSpeedMin - fSpeedMin) <> (fSpeedMin - fSpeedMin)) THEN // 转速阈值越域 / the speed threshold is out of domain
    _bCfgBad := TRUE; // 判非法 / mark illegal
END_IF
IF (nRetryMax < 0) OR (nRetryMax > 9) THEN // 重试上限越域 / the retry ceiling is out of domain
    _bCfgBad := TRUE; // 判非法 / mark illegal
END_IF
IF (tStopTo <= T#0S) OR (tGapMin <= T#0S) OR (tSpinMax <= T#0S) OR (tCloseTo <= T#0S) OR (tStableMin <= T#0S) THEN // 时间引脚非正 / a time pin is not positive
    _bCfgBad := TRUE; // 判非法 / mark illegal
END_IF
IF tSpinMax <= tGapMin THEN // 降速总窗不大于最小间隔窗，违反双窗配比（R100）/ the spin window does not exceed the gap window
    _bCfgBad := TRUE; // 判非法 / mark illegal
END_IF
IF _bCfgBad AND (NOT _bFault) THEN // 组态非法且未锁存 / illegal configuration and not yet latched
    _bFault := TRUE; // 置故障锁存 / raise the fault latch
    _eFaulC := E_DL_FbsFault.eCfgIllegal; // 故障级成因（R45 配对 bError）/ the fault cause paired with bError
    _ePhase := E_DL_FbsPhase.eFault; // 迁故障相 / migrate to the fault phase
END_IF
_nRetryUse := nRetryMax; // 重试上限直通 / the retry ceiling passes through
IF _nRetryUse < 0 THEN // 下越界 / below the floor
    _nRetryUse := 0; // 回钳到零 / clamp to zero
ELSIF _nRetryUse > 9 THEN // 上越界 / above the ceiling
    _nRetryUse := 9; // 回钳到九 / clamp to nine
END_IF

// 段 4｜中止电平优先处理：任何中间态立即双断回空闲 / segment 4, the abort level takes priority, any middle phase goes both off
IF bAbort AND (NOT _bFault) THEN // 中止且未锁存 / abort while unlatched
    _ePhase := E_DL_FbsPhase.eIdle; // 回空闲相（双断由出口派生）/ back to idle, both off by derivation
END_IF

// 段 5｜相位机：ENUM + CASE，含 ELSE 非法相位兜底（R128）/ segment 5, the phase machine with an ELSE fallback
CASE _ePhase OF
E_DL_FbsPhase.eIdle: // 空闲相：变频保持，等切换申请 / idle, the VFD holds and waits
    IF bEnable AND (NOT _bFault) AND (NOT bAbort) AND rtSwap.Q THEN // 申请沿受理 / the request edge is accepted
        _nRetry := 0; // 重试计数清零 / clear the retry count
        _ePhase := E_DL_FbsPhase.eStopVfd; // 迁停变频相 / migrate to the stop phase
    END_IF

E_DL_FbsPhase.eStopVfd: // 停变频相：等变频反馈消失 / the stop phase, the feedback drop is awaited
    IF NOT bEnable THEN // 失能 / disabled
        _ePhase := E_DL_FbsPhase.eIdle; // 回空闲相 / back to idle
    ELSIF NOT bVfdFb THEN // 变频反馈已消失 / the VFD feedback has dropped
        _ePhase := E_DL_FbsPhase.eWaitSpinDown; // 迁等降速相 / migrate to the wait phase
    ELSIF tonStop.Q THEN // 反馈消失窗耗尽 / the drop window expired
        _bFault := TRUE; // 置故障锁存 / raise the fault latch
        _eFaulC := E_DL_FbsFault.eSwapTimeout; // 故障级成因（R45 配对 bError）/ the fault cause paired with bError
        _ePhase := E_DL_FbsPhase.eFault; // 迁故障相 / migrate to the fault phase
    END_IF

E_DL_FbsPhase.eWaitSpinDown: // 等降速相：转速阈值 + 最小间隔窗 + 总窗三判（退出条件 ≥2，R98）/ the wait phase, three verdicts and at least two exit conditions
    IF NOT bEnable THEN // 失能 / disabled
        _ePhase := E_DL_FbsPhase.eIdle; // 回空闲相 / back to idle
    ELSIF tonSpin.Q THEN // 降速总窗耗尽 / the spin window expired
        _bFault := TRUE; // 置故障锁存 / raise the fault latch
        _eFaulC := E_DL_FbsFault.eSwapTimeout; // 故障级成因（R45 配对 bError）/ the fault cause paired with bError
        _ePhase := E_DL_FbsPhase.eFault; // 迁故障相 / migrate to the fault phase
    ELSIF (fSpeed <= fSpeedMin) AND tonGap.Q THEN // 转速达标且最小间隔窗已过 / the speed is low and the gap window elapsed
        _ePhase := E_DL_FbsPhase.eCloseBypass; // 迁关旁通相 / migrate to the close phase
    END_IF

E_DL_FbsPhase.eCloseBypass: // 关旁通相：出命令等反馈，失败重试 / the close phase, the command waits for the feedback with retries
    IF NOT bEnable THEN // 失能 / disabled
        _ePhase := E_DL_FbsPhase.eIdle; // 回空闲相 / back to idle
    ELSIF bBypassFb THEN // 旁通反馈确认 / the bypass feedback confirmed
        _ePhase := E_DL_FbsPhase.eRunDurance; // 迁稳定中相 / migrate to the run in phase
    ELSIF tonClose.Q THEN // 确认窗耗尽 / the confirm window expired
        IF _nRetry < _nRetryUse THEN // 重试未用尽 / retries remain
            _nRetry := _nRetry + 1; // 重试计数递增 / increment the retry count
            _ePhase := E_DL_FbsPhase.eWaitSpinDown; // 回等降速相重走间隔窗 / back to the wait phase for a fresh gap
        ELSE // 重试用尽 / retries exhausted
            _bFault := TRUE; // 置故障锁存 / raise the fault latch
            _eFaulC := E_DL_FbsFault.eRetryExhausted; // 故障级成因（R45 配对 bError）/ the fault cause paired with bError
            _ePhase := E_DL_FbsPhase.eFault; // 迁故障相 / migrate to the fault phase
        END_IF
    END_IF

E_DL_FbsPhase.eRunDurance: // 稳定中相：旁通保持，驻留稳定窗 / the run in phase, the bypass holds through the dwell window
    IF NOT bEnable THEN // 失能 / disabled
        _ePhase := E_DL_FbsPhase.eIdle; // 回空闲相 / back to idle
    ELSIF NOT bBypassFb THEN // 旁通反馈丢失 / the bypass feedback was lost
        _bFault := TRUE; // 置故障锁存 / raise the fault latch
        _eFaulC := E_DL_FbsFault.eFbLost; // 故障级成因（R45 配对 bError）/ the fault cause paired with bError
        _ePhase := E_DL_FbsPhase.eFault; // 迁故障相 / migrate to the fault phase
    ELSIF tonStable.Q THEN // 稳定驻留窗已过 / the dwell window elapsed
        _ePhase := E_DL_FbsPhase.eStable; // 迁已稳定相 / migrate to the stable phase
    END_IF

E_DL_FbsPhase.eStable: // 已稳定相：旁通运行，持续监视反馈 / the stable phase, the bypass runs with a continuous feedback watch
    IF NOT bEnable THEN // 失能 / disabled
        _ePhase := E_DL_FbsPhase.eIdle; // 回空闲相 / back to idle
    ELSIF NOT bBypassFb THEN // 旁通反馈丢失 / the bypass feedback was lost
        _bFault := TRUE; // 置故障锁存 / raise the fault latch
        _eFaulC := E_DL_FbsFault.eFbLost; // 故障级成因（R45 配对 bError）/ the fault cause paired with bError
        _ePhase := E_DL_FbsPhase.eFault; // 迁故障相 / migrate to the fault phase
    END_IF

E_DL_FbsPhase.eFault: // 故障相：双断，等复位沿 / the fault phase, both off until the reset edge
    IF NOT bEnable THEN // 失能 / disabled
        _ePhase := E_DL_FbsPhase.eIdle; // 迁未使能相 / migrate to idle
    END_IF

ELSE // 非法相位兜底（R128）/ the illegal phase fallback
    _bFault := TRUE; // 置故障锁存 / raise the fault latch
    _eFaulC := E_DL_FbsFault.ePhaseBad; // 故障级成因（R45 配对 bError）/ the fault cause paired with bError
    _ePhase := E_DL_FbsPhase.eFault; // 迁故障相 / migrate to the fault phase
END_CASE

// 段 6｜命令出口派生（互斥不变量的结构性承载）/ segment 6, the command outlets, the structural carrier of the mutual exclusion
bVfdRun := (_ePhase = E_DL_FbsPhase.eIdle) AND bEnable AND (NOT _bFault) AND (NOT bAbort); // 变频保持命令：仅空闲相派生 / the VFD hold command, derived in the idle phase only
bBypassRun := (_ePhase = E_DL_FbsPhase.eCloseBypass) OR (_ePhase = E_DL_FbsPhase.eRunDurance) OR (_ePhase = E_DL_FbsPhase.eStable); // 旁通命令：三旁通相派生 / the bypass command, derived in the three bypass phases
bBothOff := (NOT bVfdRun) AND (NOT bBypassRun); // 双断指示派生 / the both off indicator derived
nRetry := _nRetry; // 重试计数出口 / the retry count outlet

// 段 7｜统一出口 / segment 7, the unified outlet
IF _bFault THEN // 故障锁存优先 / the fault latch takes priority
    eFault := _eFaulC; // 故障级成因锁存回放（R152）/ the fault cause replayed from the latch
ELSE
    eFault := E_DL_FbsFault.eNone; // 无锁存即无成因 / no latch, no cause
END_IF
ePhase := _ePhase; // 相位出口单点映射 / single point phase outlet mapping
bError := _bFault; // 故障标志与锁存位同源 / the fault flag shares the latch source
END_FUNCTION_BLOCK

(* ---- FB_DL_FilmSpliceCurtain.st ---- *)
(*
  FB_DL_FilmSpliceCurtain  —  接膜工位光幕屏蔽序列（2 传感器模式屏蔽时序） / Film-splice station light-curtain muting sequence with two-sensor pattern
  分类 Category : DL_Device
  版本 Version  : 1.0.0
  来源 Source   : t2-8-isa182 — 安全屏蔽族深化（与 I_DL_SafetyDoor 单门接口分工：本件为光幕屏蔽时序件）
  溯源 Origin   : clean-room 实现，双传感器屏蔽模式为 ISA182 惯例公开借鉴，未复制任何源码行
  功能 Function : 1) 三相屏蔽时序：eIdle → eSeq（首传感器沿后等第二传感器沿，
                  tSeqTo 超时判）→ eMute（双传感器齐备，屏蔽承载 bMuteEn，
                  物料通过双传感器回落回 eIdle）；
                  2) 屏蔽期内光幕遮断被容忍（不置故障，屏蔽语义承载）；
                  屏蔽相滞留超 tMuteMax → 0523 锁存并退出屏蔽（安全侧）；
                  3) 非法模式：eSeq 相单传感器悬置 tSeqTo → 0522 锁存
                  （R190 归因唯一：非法模式走 0522，滞留超窗走 0523）；
                  4) 故障级：0522 屏蔽序列非法模式锁存 / 0523 屏蔽相滞留超窗
                  锁存 / 0524 组态非法（窗域）+ ELSE 兜底归并；
                  5) 信息级三码：屏蔽激活 / 屏蔽解除 / 非法模式检出（单拍沿）；
                  6) 解除式全当拍量（R240 落地），逐 BOOL 标注见段 4。
  边界 Boundary : ① 分段理由（R192）：段 0003 故障带 03A0~03FF 于 R42 用尽，
                  启用 05xx 副带续编，避开 0590~0599 判错位段；
                  ② 组态闸：tSeqTo <= 0 或 tMuteMax <= 0 → 0524 锁存；
                  ③ 安全侧：故障锁存期 bMuteEn 强制 FALSE（光幕恢复全防护）；
                  ④ 无 GVL 依赖：纯引脚输入输出，无外部变量引用，无物理 IO 地址。
  依赖 Depends  : Standard.library（TON / R_TRIG）
  码表 Error codes（Device 段 0003，窗口 0522~0524 / 0428~042A）:
    16#0003_0522 故障级：屏蔽序列非法模式锁存（单传感器悬置 tSeqTo），锁存至 bReset
    16#0003_0523 故障级：屏蔽相滞留超窗锁存（tMuteMax），锁存至 bReset
    16#0003_0524 故障级：组态非法（任一窗域非法）或相位落 ELSE 兜底（归并声明），锁存至 bReset
    16#0003_0428 信息级：屏蔽激活沿（进 eMute）
    16#0003_0429 信息级：屏蔽解除沿（回 eIdle）
    16#0003_042A 信息级：非法模式检出沿（0522 锁存拍）
  修订历史 Revision :
    2026-11-19  v1.0.0  R42 首版（批次 4 · 序号 3）
*)

TYPE E_DL_FscState :
(
    eIdle  := 0,     // 全防护：屏蔽未承载 / Full protection, muting off
    eSeq   := 10,    // 序列：等第二传感器沿 / Sequence, waiting second sensor
    eMute  := 20,    // 屏蔽：双传感器承载 / Muting, dual-sensor engaged
    eFault := 90     // 故障：非法模式或滞留锁定 / Fault, latched
);
END_TYPE

FUNCTION_BLOCK FB_DL_FilmSpliceCurtain
VAR_INPUT
    bMuteA       : BOOL := FALSE;     // 屏蔽传感器 A（当拍量）[-] / Muting sensor A, current-scan
    bMuteB       : BOOL := FALSE;     // 屏蔽传感器 B（当拍量）[-] / Muting sensor B, current-scan
    bCurtainBrk  : BOOL := FALSE;     // 光幕遮断（当拍量，TRUE = 遮断）[-] / Light curtain broken flag
    tSeqTo       : TIME := T#2S;      // 序列第二传感器等待窗 [ms]，域 > 0 / Sequence second-sensor window
    tMuteMax     : TIME := T#10S;     // 屏蔽最大承载窗 [ms]，域 > 0 / Maximum muting window
    bReset       : BOOL := FALSE;     // 复位，上升沿清故障锁存 / Reset edge clears fault latch
END_VAR
VAR_OUTPUT
    eState       : E_DL_FscState;     // 状态出口，段尾单点映射 / State outlet
    bMuteEn      : BOOL;              // 屏蔽承载输出（eMute 相电平）[-] / Muting engage output
    bCurtainSafe : BOOL;              // 光幕安全出口（遮断且非屏蔽 → FALSE）[-] / Curtain safety outlet
    bError       : BOOL;              // 故障锁存标志 / Fault latch flag
    nErrId       : UDINT;             // 事件码，0 = 无事件 / Event code
END_VAR
VAR
    tonSeqTo     : TON;               // 序列等待窗（单相独占），无条件刷新 / Sequence window timer
    tonMuteMax   : TON;               // 屏蔽承载窗（单相独占），无条件刷新 / Muting window timer
    rtMuteA      : R_TRIG;            // 传感器 A 沿实例，无条件刷新 / Sensor A edge instance
    rtMuteB      : R_TRIG;            // 传感器 B 沿实例，无条件刷新 / Sensor B edge instance
    rtReset      : R_TRIG;            // 复位沿实例，无条件刷新 / Reset edge instance
    _eState      : E_DL_FscState := E_DL_FscState.eIdle;  // 内部相位（CASE 唯一写入目标）/ Internal phase
    _bFault      : BOOL;              // 故障锁存位（锁存量）/ Latched fault bit
    _uFault      : UDINT;             // 故障码锁存（锁存量）/ Latched fault code
    _uInfo       : UDINT;             // 信息码，每拍重算 / Transient info code
END_VAR

(* —— 段 0：定时器与沿实例无条件周期刷新（禁置于 IF/CASE 内） —— *)
rtMuteA(CLK := bMuteA);              // 传感器 A 沿（每拍必调）
rtMuteB(CLK := bMuteB);              // 传感器 B 沿（每拍必调）
rtReset(CLK := bReset);              // 复位沿（每拍必调）
tonSeqTo(IN := (_eState = E_DL_FscState.eSeq), PT := tSeqTo);        // 序列窗（单相独占）
tonMuteMax(IN := (_eState = E_DL_FscState.eMute), PT := tMuteMax);   // 屏蔽窗（单相独占）

(* —— 段 1：单拍量预清零（锁存量 _bFault/_uFault 不入清单，禁同拍抹除） —— *)
_uInfo := 16#0000_0000;             // 信息码每拍重算
bMuteEn := FALSE;                   // 屏蔽输出缺省 FALSE（安全侧）
bCurtainSafe := FALSE;              // 光幕安全出口缺省 FALSE（安全侧）
nErrId := 16#0000_0000;             // 事件码缺省无事件

(* —— 段 2：复位沿 + 组态域闸（判据当拍量） —— *)
IF rtReset.Q THEN                   // rtReset.Q = 当拍量
    _bFault := FALSE;               // 清故障锁存位
    _uFault := 16#0000_0000;        // 清故障锁存码
END_IF
IF (TIME_TO_DINT(tSeqTo) <= 0) OR (TIME_TO_DINT(tMuteMax) <= 0) THEN
    _uFault := 16#0003_0524;        // 故障级：组态非法
    _bFault := TRUE;                // 故障标志与码位配对（R45）
END_IF

(* —— 段 3：非法模式与滞留超窗锁存（判据当拍量/单相独占 TON） —— *)
IF (NOT _bFault) AND tonSeqTo.Q THEN
    _uFault := 16#0003_0522;        // 故障级：非法模式（单传感器悬置）
    _bFault := TRUE;
    _uInfo := 16#0003_042A;         // 信息级：非法模式检出沿
END_IF
IF (NOT _bFault) AND tonMuteMax.Q THEN
    _uFault := 16#0003_0523;        // 故障级：屏蔽相滞留超窗
    _bFault := TRUE;
END_IF

(* —— 段 4：故障解除式（R240 落地，逐 BOOL 标注）：
     rtReset.Q = 当拍量；NOT bMuteA = 当拍量；NOT bMuteB = 当拍量；
     NOT bCurtainBrk = 当拍量。均不含锁存量（_bFault/_uFault），
     解除边真实可达（双传感器回落 + 光幕恢复 + 复位沿）。 —— *)
IF rtReset.Q AND (NOT bMuteA) AND (NOT bMuteB) AND (NOT bCurtainBrk) THEN
    _bFault := FALSE;               // 清故障锁存位（锁存量，仅此当拍量解除沿可清）
    _uFault := 16#0000_0000;        // 清故障锁存码（锁存量，仅本当拍量解除沿可清）
    IF _eState = E_DL_FscState.eFault THEN
        _eState := E_DL_FscState.eIdle;     // 故障相迁出：回全防护
    END_IF
END_IF

(* —— 段 5：相位机（CASE 全覆盖 + ELSE 兜底） —— *)
CASE _eState OF

E_DL_FscState.eIdle:
    IF rtMuteA.Q OR rtMuteB.Q THEN  // 任一传感器沿：进序列相
        _eState := E_DL_FscState.eSeq;
    END_IF

E_DL_FscState.eSeq:
    IF (rtMuteA.Q AND bMuteB) OR (rtMuteB.Q AND bMuteA) THEN
        _uInfo := 16#0003_0428;     // 信息级：屏蔽激活沿（第二传感器齐备拍）
        _eState := E_DL_FscState.eMute;     // 进屏蔽相
    END_IF
    (* 非法模式迁出在段 3 承载 *)

E_DL_FscState.eMute:
    IF (NOT bMuteA) AND (NOT bMuteB) THEN   // 双传感器回落：物料通过
        _uInfo := 16#0003_0429;     // 信息级：屏蔽解除沿
        _eState := E_DL_FscState.eIdle;     // 回全防护相
    END_IF
    (* 滞留超窗迁出在段 3 承载 *)

E_DL_FscState.eFault:
    ;                               // 故障相：屏蔽强制断，等解除沿（段 4 承载迁出）

ELSE
    _uFault := 16#0003_0524;        // 故障级：非法相位兜底（归并组态码，码表声明）
    _bFault := TRUE;
    _eState := E_DL_FscState.eFault;    // 强制回故障相

END_CASE

(* —— 段 6：出口单点映射（名实同源；锁存码回放，禁同拍抹除） —— *)
IF _eState = E_DL_FscState.eMute THEN
    bMuteEn := TRUE;                // 屏蔽承载（相电平）
    bCurtainSafe := TRUE;           // 屏蔽期光幕遮断被容忍（安全出口保持 TRUE）
ELSIF bCurtainBrk THEN
    bCurtainSafe := FALSE;          // 非屏蔽期遮断：安全出口 FALSE（全防护语义）
ELSE
    bCurtainSafe := TRUE;           // 非屏蔽期未遮断：安全出口 TRUE
END_IF
IF _bFault THEN
    nErrId := _uFault;              // 故障锁存码回放
    bMuteEn := FALSE;               // 故障相屏蔽强制 FALSE（安全侧，③声明）
    bCurtainSafe := NOT bCurtainBrk;    // 故障相光幕语义保持全防护（遮断即 FALSE）
ELSE
    nErrId := _uInfo;               // 信息码
END_IF
bError := _bFault;                  // 故障标志与锁存位同源
eState := _eState;                  // 状态出口单点映射

END_FUNCTION_BLOCK

(* ---- FB_DL_FilterDpMonitor.st ---- *)
//==============================================================================
// 功能块：FB_DL_FilterDpMonitor ｜ 中文名称：过滤器压差寿命监视
// 所属子库：DL_Device ｜ 版本：v1.0.0 ｜ 兼容：CODESYS V3.5+ / TwinCAT 3 / 汇川 InoProShop
// 功能描述：过滤器压差趋势监视与滤芯更换预警——压差实测 + 趋势窗斜率
//           [kPa/h]，按更换预警/堵塞报警双阈值映射 NE107 健康态
//           （eOk / eMaintenanceReq / eOutOfSpec），eOutOfSpec 锁存需手动复位。
// 开源溯源 (Origin)：道莅 clean-room 防御性实现
// 单位表：p_d[kPa] / 趋势斜率[kPa/h] / 阈值[kPa] / 趋势窗[ms] / 健康态[—]
// 错误码表：16#0003_0182 信息级（负压差，传感器接反疑似，按 0 处理，不置
//           bError）/ 16#0003_0183 预留禁用（不得挪用）/ 16#0003_0354
//           故障级（阈值倒置或压差非有限，置 bError，保持末次有效健康态）/
//           16#0003_0355 预留禁用（不得挪用）/ 16#0003_0356 故障级兜底
//           （置 bError，本件无状态机，保留给扩展误用拦截）
// 状态机：N/A（阈值映射 + 锁存为电平逻辑，无相位状态机；健康态降级锁存
//           由 bOosLatch 保持量承担）
// 边界行为：① fDpAlarmKpa <= fDpChangeKpa → 故障 0354（阈值倒置）；② 压差
//           非有限 → 故障 0354 复用（R90）+ 保持末次有效健康态（不静默塞
//           eOk）；③ 负压差（传感器接反疑似）→ 信息 0182 + 按 0 处理；
//           ④ 趋势窗斜率 = 窗均值差 / 窗时长[h]，窗时长非法（<= 0）→ 斜率
//           冻结 0（防除零）；⑤ eOutOfSpec 锁存，仅 bReset 清除。
// 依赖纪律：Level 1 → Level 0 组合调用合法——趋势窗均值组合调用
//           FB_DL_SignalStatistics（DL_MathData，接口已核实：fIn/bSample/
//           nWindow/bClear → fMean/fMin/fMax/fRange/fVariance），头注释
//           依赖清单声明；斜率除法在本件内联（时间维度归一属监视语义，
//           非统计算法复制）。
// 修订历史：v1.0.0 2026-11-17 首版（R23 派单 · ROADMAP 公用工程 P1 §394 + T2-8 NE107 次源）
//==============================================================================

FUNCTION_BLOCK FB_DL_FilterDpMonitor
VAR_INPUT
    fDpKpa       : LREAL;                    // 压差实测 [千帕] / Measured differential pressure [kPa]
    fDpChangeKpa : LREAL := 0.8;             // 更换预警阈值 [千帕] / Replace-hint threshold [kPa]
    fDpAlarmKpa  : LREAL := 1.5;             // 堵塞报警阈值 [千帕]，须 > 预警阈值 / Clog-alarm threshold [kPa], must exceed the hint threshold
    tTrendWindow : TIME  := T#1H;            // 趋势窗时长 [ms] / Trend window duration [ms]
    bReset       : BOOL;                     // 手动复位 [—]，清除 eOutOfSpec 锁存 / Manual reset, clears the eOutOfSpec latch
END_VAR
VAR_OUTPUT
    eHealth      : E_DL_Ne107Status;         // 健康态 [—]，引用属主枚举（只引用不重声明，R70） / Health status, owner enum referenced, not redeclared
    fDpTrendKpaH : LREAL;                    // 趋势斜率 [千帕/小时] / Trend slope [kPa/h]
    bReplaceHint : BOOL;                     // 更换预警 [—] / Replace hint
    eErr         : UDINT;                    // 错误码，0 = 无错 / Error code, 0 = no error
    bError       : BOOL;                     // 故障级标志，仅故障级错误置位 / Fault-class flag, set only on fault-level codes
    bValid       : BOOL;                     // 输出可用标志 / Outputs usable flag
END_VAR
VAR
    fbStats      : FB_DL_SignalStatistics;   // 趋势窗统计器（Level 0 组合调用） / Trend-window statistics FB, Level 0 composition
    fbWin        : TON;                      // 趋势窗计时，段 6 无条件刷新 [ms] / Trend window timer
    rtWinTick    : R_TRIG;                   // 窗满上升沿（快照单发），段 6 无条件刷新 / Window-full rising edge, one-shot snapshot
    _eHealthAcc  : E_DL_Ne107Status := E_DL_Ne107Status.eUnknown; // 末次有效健康态保持量 / Held last valid health status
    _bOosLatch   : BOOL;                     // eOutOfSpec 锁存（bReset 清除） / eOutOfSpec latch, cleared by bReset
    _fMeanPrev   : REAL;                     // 上一窗均值快照 [千帕] / Previous window-mean snapshot [kPa]
    _fWinHours   : LREAL;                    // 趋势窗时长换算 [小时] / Trend window duration [h]
    _fDpEff      : LREAL;                    // 防御后的生效压差 [千帕] / Effective defended pressure [kPa]
    _bInit       : BOOL := FALSE;            // 首扫标志，初值 FALSE 取非判定 / First-scan flag, tested negated
    _bThreshBad  : BOOL;                    // 阈值倒置锁存 / Threshold inversion latch
    _bFiniteBad  : BOOL;                    // 压差非有限锁存 / Non-finite pressure latch
    _bNegDp      : BOOL;                     // 负压差当拍标志 / Negative pressure flag of this scan
END_VAR
VAR CONSTANT
    DL_FD_INF     : LREAL := 1.7976931348623157E308; // LREAL 幅值上限 / LREAL magnitude ceiling
    DL_FD_ZERO    : LREAL := 0.0;          // 压差物理下界 [千帕] / Pressure physical floor [kPa]
    DL_FD_H_PER_MS: LREAL := 2.77777777777778E-7; // 毫秒 → 小时换算系数 [h/ms]，1/3600000 / Millisecond-to-hour factor [h/ms]
    DL_FD_STATS_N : INT   := 32;           // 统计窗口长度 [样本] / Statistics window length [samples]
END_VAR

(*------------------------------------------------------------------------------
 * 段 1｜每拍预置：输出先算后出，单拍标志预清零
 *      Outputs computed per scan, one-shot flags pre-cleared
 *-----------------------------------------------------------------------------*)
eHealth      := E_DL_Ne107Status.eUnknown; // 健康态预置未知 / Health preset unknown
fDpTrendKpaH := 0.0;                       // 趋势斜率预置零 / Trend slope preset zero
bReplaceHint := FALSE;                     // 更换预警预清零 / Replace hint pre-cleared
eErr         := 16#0000_0000;              // 错误码每拍重算 / Error code recomputed
bError       := FALSE;                     // 故障标志每拍重算 / Fault flag recomputed
bValid       := FALSE;                     // 可用标志每拍重算 / Usable flag recomputed
_bNegDp      := FALSE;                     // 负压差标志预清零 / Negative flag pre-cleared

(*------------------------------------------------------------------------------
 * 段 2｜首扫初始化
 *      First-scan initialisation
 *-----------------------------------------------------------------------------*)
IF NOT _bInit THEN
    _eHealthAcc := E_DL_Ne107Status.eOk;   // 末次有效健康态起步正常 / Held health starts OK
    _fMeanPrev  := 0.0;                    // 均值快照清零 / Mean snapshot cleared
    _bOosLatch  := FALSE;                  // 超规格锁存清零 / OOS latch cleared
    _bInit      := TRUE;                   // 首扫只做一次 / The first scan runs once
END_IF

(*------------------------------------------------------------------------------
 * 段 3｜组态与输入防御闸：阈值倒置 / 非有限 → 0354（保持末次健康态）
 *      Configuration and input defense gate, last valid health held
 *-----------------------------------------------------------------------------*)
IF fDpAlarmKpa <= fDpChangeKpa THEN
    _bThreshBad := TRUE;                   // 阈值倒置锁存 / Threshold inversion latched
END_IF
IF (fDpKpa <> fDpKpa) OR (ABS(fDpKpa) > DL_FD_INF) THEN
    _bFiniteBad := TRUE;                   // 压差非有限锁存 / Non-finite pressure latched
END_IF

(*------------------------------------------------------------------------------
 * 段 4｜负压差防御：传感器接反疑似，按 0 处理并声明
 *      Negative pressure defense, treated as zero with a notice
 *-----------------------------------------------------------------------------*)
_fDpEff := fDpKpa;                          // 生效压差先取原值 / Effective pressure starts as-is
IF (NOT _bFiniteBad) AND (fDpKpa < DL_FD_ZERO) THEN
    _bNegDp := TRUE;                        // 负压差当拍成立 / Negative pressure active this scan
    _fDpEff := 0.0;                         // 负压差按 0 处理 / Negative pressure treated as zero
END_IF

(*------------------------------------------------------------------------------
 * 段 5｜趋势组合调用与窗计时无条件刷新（R40：CASE 之外每拍必调）
 *      Trend composition and window timing refreshed unconditionally
 *-----------------------------------------------------------------------------*)
fbStats(fIn := LREAL_TO_REAL(_fDpEff), bSample := TRUE, nWindow := DL_FD_STATS_N); // 统计器每拍采样（标准类型转换，零方言） / Statistics FB sampled every scan, standard type conversion
fbWin(IN := TRUE, PT := tTrendWindow);     // 趋势窗连续计时 / Trend window timing continuous
rtWinTick(CLK := fbWin.Q);                 // 窗满上升沿 / Window-full edge
_fWinHours := TIME_TO_DINT(tTrendWindow) * DL_FD_H_PER_MS; // 窗时长换算 [小时] / Window duration converted [h]
IF rtWinTick.Q AND (_fWinHours > 0.0) THEN
    fDpTrendKpaH := (fbStats.fMean - _fMeanPrev) / _fWinHours; // 趋势斜率 [千帕/小时]，分母已闸 / Trend slope, denominator gated
    _fMeanPrev := fbStats.fMean;           // 快照推进 / Snapshot advanced
ELSIF _fWinHours <= 0.0 THEN
    fDpTrendKpaH := 0.0;                   // 窗时长非法：斜率冻结（防除零） / Illegal duration, slope frozen, divide-by-zero guarded
END_IF

(*------------------------------------------------------------------------------
 * 段 6｜阈值映射与降级锁存（eOutOfSpec 需手动复位才回 eOk）
 *      Threshold mapping and the degradation latch
 *-----------------------------------------------------------------------------*)
IF (NOT _bThreshBad) AND (NOT _bFiniteBad) THEN
    bReplaceHint := (_fDpEff >= fDpChangeKpa); // 生效压差达预警阈值 / Effective pressure at the hint threshold
    IF _fDpEff >= fDpAlarmKpa THEN
        _bOosLatch := TRUE;                // 达报警阈值，锁存超规格 / At the alarm threshold, OOS latched
    END_IF
    IF _bOosLatch THEN
        _eHealthAcc := E_DL_Ne107Status.eOutOfSpec; // 锁存期保持超规格 / OOS held during the latch
    ELSIF bReplaceHint THEN
        _eHealthAcc := E_DL_Ne107Status.eMaintenanceReq; // 预警期维护请求 / Maintenance required during the hint
    ELSE
        _eHealthAcc := E_DL_Ne107Status.eOk; // 正常 / OK
    END_IF
END_IF
IF bReset THEN
    _bOosLatch := FALSE;                   // 手动复位清锁存 / Manual reset clears the latch
END_IF

(*------------------------------------------------------------------------------
 * 段 7｜输出与码位出口
 *      Outputs and the code outlet
 *-----------------------------------------------------------------------------*)
eHealth := _eHealthAcc;                    // 健康态出口（故障期保持末次有效值） / Health outlet, last valid value held on fault
IF _bThreshBad OR _bFiniteBad THEN
    eErr   := 16#0003_0354;                // 故障级：阈值倒置或非有限（R90 复用） / Fault: threshold inversion or non-finite, code reused
    bError := TRUE;                        // 置故障标志（R45 配对） / Raise the fault flag
    bValid := FALSE;                       // 输出不可用 / Outputs unusable
ELSE
    IF _bNegDp THEN
        eErr := 16#0003_0182;              // 信息级：负压差按 0 处理（不置 bError） / Info: negative pressure treated as zero, no fault flag
    END_IF
    bValid := TRUE;                        // 输出可用 / Outputs usable
END_IF
END_FUNCTION_BLOCK
